(* Logix 5000 project; controller TFF vendor 1 type 14 code 107 rev 34.11; software revision 34.03; part 4 of 36 *)

        BufferEvents[140] := '07242026,07:35:58.6,700003,0.0,1.00000000', BufferEvents[141] := '07242026,07:35:58.7,1300205,2.00000000,4.00000000', BufferEvents[142] := '07242026,07:35:58.7,1300405,2.00000000,4.00000000', BufferEvents[143] := '07242026,07:35:58.7,1300505,2.00000000,4.00000000', BufferEvents[144] := '07242026,07:35:58.7,1300605,2.00000000,4.00000000', BufferEvents[145] := '07242026,07:35:58.7,1301105,2.00000000,4.00000000', BufferEvents[146] := '07242026,07:35:58.7,1301205,2.00000000,4.00000000', BufferEvents[147] := '07242026,07:35:58.7,1301305,2.00000000,4.00000000', BufferEvents[148] := '07242026,07:35:58.7,1301405,2.00000000,4.00000000', BufferEvents[149] := '07242026,07:35:58.8,2500101,0.0,1.00000000', BufferEvents[150] := '07242026,07:35:58.8,2500401,0.0,1.00000000', BufferEvents[151] := '07242026,07:35:58.8,2500801,1.00000000,0.0', BufferEvents[152] := '07242026,07:35:58.8,2501901,0.0,1.00000000', BufferEvents[153] := '07242026,08:54:51.3,305106,1.00000000,0.0', BufferEvents[154] := '07242026,08:55:09.5,305206,1.00000000,0.0', BufferEvents[155] := '07242026,08:56:06.6,305006,1.00000000,0.0', BufferEvents[156] := '07242026,09:12:34.6,300107,0.0,1.00000000', BufferEvents[157] := '07242026,09:14:51.8,700003,1.00000000,0.0', BufferEvents[158] := '07242026,09:14:51.8,300106,1.00000000,0.0', BufferEvents[159] := '07242026,09:14:51.8,300607,0.0,1.00000000', BufferEvents[160] := '07242026,09:14:51.8,300707,0.0,1.00000000', BufferEvents[161] := '07242026,09:14:51.9,305006,0.0,1.00000000', BufferEvents[162] := '07242026,09:14:51.9,305106,0.0,1.00000000', BufferEvents[163] := '07242026,09:14:51.9,305206,0.0,1.00000000', BufferEvents[164] := '07242026,09:14:51.9,1600003,1.00000000,0.0', BufferEvents[165] := '07242026,09:14:51.9,1300205,4.00000000,2.00000000', BufferEvents[166] := '07242026,09:14:51.9,1300405,4.00000000,2.00000000', BufferEvents[167] := '07242026,09:14:51.9,1300505,4.00000000,2.00000000', BufferEvents[168] := '07242026,09:14:51.9,1300605,4.00000000,2.00000000', BufferEvents[169] := '07242026,09:14:51.9,1301105,4.00000000,2.00000000', BufferEvents[170] := '07242026,09:14:51.9,1301205,4.00000000,2.00000000', BufferEvents[171] := '07242026,09:14:51.9,1301305,4.00000000,2.00000000', BufferEvents[172] := '07242026,09:14:51.9,1301405,4.00000000,2.00000000', BufferEvents[173] := '07242026,09:14:52.0,2500101,1.00000000,0.0', BufferEvents[174] := '07242026,09:14:52.0,2500401,1.00000000,0.0', BufferEvents[175] := '07242026,09:14:52.0,2500801,0.0,1.00000000', BufferEvents[176] := '07242026,09:14:52.0,2501901,1.00000000,0.0', BufferEvents[177] := '07242026,09:14:52.9,306806,1.00000000,0.0', BufferEvents[178] := '07242026,09:14:55.0,1600003,0.0,1.00000000', BufferEvents[179] := '07242026,09:14:56.8,305506,1.00000000,0.0', BufferEvents[180] := '07242026,09:14:56.8,305706,1.00000000,0.0', BufferEvents[181] := '07242026,09:14:56.8,306906,1.00000000,0.0', BufferEvents[182] := '07242026,09:14:56.8,307106,1.00000000,0.0', BufferEvents[183] := '07242026,09:14:56.8,307306,1.00000000,0.0', BufferEvents[184] := '07242026,09:14:56.8,307506,1.00000000,0.0', BufferEvents[185] := '07242026,09:15:07.7,300106,0.0,1.00000000', BufferEvents[186] := '07242026,09:15:07.7,306806,0.0,1.00000000', BufferEvents[187] := '07242026,09:15:07.7,300107,1.00000000,0.0', BufferEvents[188] := '07242026,09:15:07.7,300607,1.00000000,0.0', BufferEvents[189] := '07242026,09:15:07.7,300707,1.00000000,0.0', BufferEvents[190] := '07242026,09:15:07.8,300306,1.00000000,0.0', BufferEvents[191] := '07242026,09:15:09.7,300006,1.00000000,0.0', BufferEvents[192] := '07242026,09:19:10.3,305506,0.0,1.00000000', BufferEvents[193] := '07242026,09:19:10.3,305706,0.0,1.00000000', BufferEvents[194] := '07242026,09:19:10.3,307106,0.0,1.00000000', BufferEvents[195] := '07242026,09:19:10.3,307306,0.0,1.00000000', BufferEvents[196] := '07242026,09:19:10.3,307506,0.0,1.00000000', BufferEvents[197] := '07242026,09:19:10.3,1600003,1.00000000,0.0', BufferEvents[198] := '07242026,09:19:13.4,1600003,0.0,1.00000000', BufferEvents[199] := '07242026,09:19:17.6,300306,0.0,1.00000000',
        BufferEvents[200] := '07242026,09:19:18.6,300006,0.0,1.00000000', BufferEvents[201] := '07242026,09:19:35.6,306906,0.0,1.00000000', BufferEvents[202] := '07242026,09:19:36.6,300806,1.00000000,0.0', BufferEvents[203] := '07242026,09:19:36.6,300906,1.00000000,0.0', BufferEvents[204] := '07242026,09:19:37.7,301006,1.00000000,0.0', BufferEvents[205] := '07242026,09:19:39.5,300806,0.0,1.00000000', BufferEvents[206] := '07242026,09:19:39.5,300906,0.0,1.00000000', BufferEvents[207] := '07242026,09:19:39.5,301006,0.0,1.00000000', BufferEvents[208] := '07242026,09:19:39.5,1600003,1.00000000,0.0', BufferEvents[209] := '07242026,09:19:42.6,1600003,0.0,1.00000000', BufferEvents[210] := '07242026,10:57:37.4,700003,0.0,1.00000000', BufferEvents[211] := '07242026,10:57:37.5,1300205,2.00000000,4.00000000', BufferEvents[212] := '07242026,10:57:37.5,1300405,2.00000000,4.00000000', BufferEvents[213] := '07242026,10:57:37.5,1300505,2.00000000,4.00000000', BufferEvents[214] := '07242026,10:57:37.5,1300605,2.00000000,4.00000000', BufferEvents[215] := '07242026,10:57:37.5,1301105,2.00000000,4.00000000', BufferEvents[216] := '07242026,10:57:37.5,1301205,2.00000000,4.00000000', BufferEvents[217] := '07242026,10:57:37.5,1301305,2.00000000,4.00000000', BufferEvents[218] := '07242026,10:57:37.5,1301405,2.00000000,4.00000000', BufferEvents[219] := '07242026,10:57:37.6,2500101,0.0,1.00000000', BufferEvents[220] := '07242026,10:57:37.6,2500401,0.0,1.00000000', BufferEvents[221] := '07242026,10:57:37.6,2500801,1.00000000,0.0', BufferEvents[222] := '07242026,10:57:37.6,2501901,0.0,1.00000000', BufferEvents[223] := '07242026,10:57:44.5,900103,1.00000000,0.0', BufferEvents[224] := '07242026,10:57:48.7,500106,30.0000000,0.0', BufferEvents[225] := '07242026,10:57:54.2,900101,1.00000000,0.0', BufferEvents[226] := '07242026,10:57:54.2,500128,1.00000000,0.0', BufferEvents[227] := '07242026,10:58:25.0,500128,0.0,1.00000000', BufferEvents[228] := '07242026,10:58:25.0,500126,1.00000000,0.0', BufferEvents[229] := '07242026,11:03:15.0,900101,0.0,1.00000000', BufferEvents[230] := '07242026,11:03:15.0,500126,0.0,1.00000000', BufferEvents[231] := '07242026,11:03:21.9,500106,0.0,30.0000000', BufferEvents[232] := '07242026,11:03:46.9,900103,0.0,1.00000000', BufferEvents[233] := '07242026,11:05:12.4,1700011,0.0,1.00000000', BufferEvents[234] := '07242026,11:05:12.5,1700003,1.00000000,0.0', BufferEvents[235] := '07242026,11:05:13.6,2600007,1.00000000,0.0', BufferEvents[236] := '07242026,11:05:13.6,2600007,0.0,1.00000000', BufferEvents[237] := '07242026,11:05:13.8,700005,10.0000000,0.0', BufferEvents[238] := '07242026,11:05:13.9,700301,1.00000000,0.0', BufferEvents[239] := '07242026,11:05:13.9,700302,0.0,1.00000000', BufferEvents[240] := '07242026,11:05:14.1,1301205,4.00000000,2.00000000', BufferEvents[241] := '07242026,11:05:14.1,1301305,4.00000000,2.00000000', BufferEvents[242] := '07242026,11:05:14.2,2502801,1.00000000,0.0', BufferEvents[243] := '07242026,11:05:14.2,1301205,2.00000000,4.00000000', BufferEvents[244] := '07242026,11:05:14.3,2502801,0.0,1.00000000', BufferEvents[245] := '07242026,11:05:14.3,2300001,1.00000000,0.0', BufferEvents[246] := '07242026,11:05:14.3,1301305,2.00000000,4.00000000', BufferEvents[247] := '07242026,11:05:14.4,2300003,1.00000000,0.0', BufferEvents[248] := '07242026,11:05:14.5,800301,1.00000000,0.0', BufferEvents[249] := '07242026,11:05:15.4,2300001,0.0,1.00000000', BufferEvents[250] := '07242026,11:05:15.5,2300003,0.0,1.00000000', DefaultOnComplete := 1);   // CCP System Data
   CCPSystem_Storage : CCPSystem_Storage[6] := ([0].Download := 1, [0].TestAction := 1, [0].State := 3, [0].Language := 1, [0].EndPointer := 34, [0].Machine := 'Mobius FlexReady', [0].Created := '03/13/2018 4:36:30 AM', [0].Originator := 'Smart', [0].OperationName := 'c:\\millipore\\CCPRecipeFiles\\SmartXMO_00.02.opn', [0].ConfigFile := 'XMO4.cfg', [0].StateWatchDog.PRE := 300000, [1].Download := 1, [1].TestAction := 1, [1].State := 3, [1].Language := 1, [1].EndPointer := 1, [1].Machine := 'Mobius FlexReady', [1].Created := '08/06/2019 8:22:36 AM', [1].Originator := 'test', [1].ConfigFile := 'TF3S.cfg', [1].StateWatchDog.PRE := 300000, [2].Download := 1, [2].TestAction := 1, [2].State := 3, [2].Language := 1, [2].EndPointer := 5, [2].Machine := 'Mobius FlexReady', [2].Created := '02/20/2018 2:20:36 AM', [2].Originator := 'QSP', [2].ConfigFile := 'MASTER_CFG--XMO4.cfg', [2].StateWatchDog.PRE := 300000, [3].Download := 1, [3].OperationDownloadFlag := 1, [3].TestAction := 1, [3].State := 3, [3].Language := 1, [3].EndPointer := 9, [3].Machine := 'Mobius FlexReady', [3].Created := '01/18/2018 5:35:26 AM', [3].Originator := 'ccc', [3].OperationName := 'c:\\millipore\\CCPRecipeFiles\\Untitled2_00.02.opn', [3].ConfigFile := 'MASTER_CFG--XMO4.cfg', [3].StateWatchDog.PRE := 300000, [4].Download := 1, [4].TestAction := 1, [4].State := 3, [4].Language := 1, [4].EndPointer := 9, [4].Machine := 'Mobius FlexReady', [4].Created := '01/18/2018 5:35:26 AM', [4].Originator := 'ccc', [4].ConfigFile := 'MASTER_CFG--XMO4.cfg', [4].StateWatchDog.PRE := 300000, [5].Download := 1, [5].OperationDownloadFlag := 1, [5].TestAction := 1, [5].State := 3, [5].Language := 1, [5].EndPointer := 9, [5].Machine := 'Mobius FlexReady',
        [5].Created := '01/18/2018 5:35:26 AM', [5].Originator := 'ccc', [5].OperationName := 'c:\\millipore\\CCPRecipeFiles\\Untitled2_00.02.opn', [5].ConfigFile := 'MASTER_CFG--XMO4.cfg', [5].StateWatchDog.PRE := 300000);
   ChartMark : ChartMark := (Out := 1);   // Chart Mark
   Concentration : Concentration := (VCF := 1.0, CB := 15.9, Conc_Init := 15.9, Conc_Final := 30.0, Final_Conc_Volume_Reached := 1, Final_Conc_Volume_DownTimer.PRE := 10000, Final_Conc_Volume_UpTimer.PRE := 1000, Final_Conc_Volume_UpTimer.ACC := 1015, Final_Conc_Volume_UpTimer.EN := 1, Final_Conc_Volume_UpTimer.DN := 1, Final_Conc_Protein_DownTimer.PRE := 10000, Final_Conc_Protein_DownTimer.ACC := 10089, Final_Conc_Protein_DownTimer.EN := 1, Final_Conc_Protein_DownTimer.DN := 1, Final_Conc_Protein_UpTimer.PRE := 1000, LogConcTimer.PRE := 3000);
   ControlLoop : ControlLoop[20] := ([0].RampTimer.PRE := 3600000, [0].StableTimer.PRE := 5000, [0].PIDTimer.PRE := 250, [0].PIDTimer.ACC := 100, [0].PIDTimer.EN := 1, [0].PIDTimer.TT := 1, [0].PID.CTL := 25199488, [0].PID.MO := 1, [0].PID.PE := 1, [0].PID.INI := 1, [0].PID.DVPA := 1, [0].PID.PVLA := 1, [0].PID.PVHA := 1, [0].PID.SP := 66.66666, [0].PID.KP := 0.5, [0].PID.KI := 0.1, [0].PID.MAXS := 200.0, [0].PID.SO := 10.0, [0].PID.MAXO := 100.0, [0].PID.MINO := 10.0, [0].PID.UPD := 0.25, [0].PID.ERR := 66.66666, [0].PID.OUT := 10.0, [0].PID.MAXI := 200.0, [0].PID.TIE := 10.0, [0].PID.MAXCV := 100.0, [0].PID.MAXTIE := 100.0, [0].PID.DATA[0] := -6.666666, [0].PID.DATA[3] := 66.66666, [0].PID.DATA[4] := 66.66666, [0].PID.DATA[5] := 0.5, [0].PID.DATA[6] := 1.0, [0].PID.DATA[7] := 4.0, [0].PID.DATA[8] := 0.5, [0].PID.DATA[9] := 0.1, [0].PID.DATA[11] := 0.5, [0].PID.DATA[12] := 0.08333334, [0].PID.DATA[15] := 1.0, [0].PID.DATA[16] := 1.0, [1].Tag := 'FIC01', [1].Desc := 'Feed Pump Control Loop', [1].LoopCfg := 1, [1].ManualEGU := '%', [1].Auto1EGU := 'LPM', [1].Auto2EGU := 'Bar', [1].Manual := 1, [1].RampEnable := 1, [1].PIDEnable := 1, [1].ManualOSR := 1, [1].PVAuto2 := 3.9859235, [1].SPAuto := 10.0, [1].SPAuto1 := 10.0, [1].SPAuto2 := 1.0, [1].RangeMax := 100.0, [1].RampRate := 1.0, [1].RampRateSave := 1.0, [1].Deadband := 10.0, [1].DBLO := 9.0, [1].DBHI := 11.0, [1].RampTimer.PRE := 3600000,
        [1].StableTimer.PRE := 10000, [1].StableTime := 10, [1].PIDTimer.PRE := 250, [1].CycleTimer.PRE := 2000, [1].PID.CTL := -2080341120, [1].PID.EN := 1, [1].PID.SWM := 1, [1].PID.INI := 1, [1].PID.DVPA := 1, [1].PID.PVLA := 1, [1].PID.PVHA := 1, [1].PID.SP := 10.0, [1].PID.KP := 0.1, [1].PID.KI := 0.2, [1].PID.MAXS := 48.0, [1].PID.DB := 0.01, [1].PID.MAXO := 100.0, [1].PID.UPD := 0.25, [1].PID.ERR := 10.0, [1].PID.MAXI := 48.0, [1].PID.MAXCV := 100.0, [1].PID.MAXTIE := 48.0, [1].PID.DATA[0] := -2.0833333, [1].PID.DATA[3] := 10.0, [1].PID.DATA[4] := 10.0, [1].PID.DATA[5] := 2.0833333, [1].PID.DATA[6] := 1.0, [1].PID.DATA[7] := 4.0, [1].PID.DATA[8] := 0.1, [1].PID.DATA[9] := 0.2, [1].PID.DATA[11] := 0.1, [1].PID.DATA[12] := 0.2, [1].PID.DATA[15] := 1.0, [1].PID.DATA[16] := 2.0833333, [1].KP[0] := 100.0, [1].KP[1] := 100.0, [1].KI[0] := 200.0, [1].KI[1] := 200.0, [1].DB[0] := 0.01, [1].Auto1Cfg := 1, [1].Auto2Cfg := 1, [1].Auto1PVCfg := 42, [1].Auto2PVCfg := 40, [1].Auto1RangeMax := 48.0, [1].Auto2RangeMax := 87.0, [1].OutputAddress := 2, [2].Tag := 'LIC01', [2].Desc := 'Level Control Loop', [2].LoopCfg := 1, [2].ManualEGU := '%', [2].Auto1EGU := 'L', [2].Interlock := 1, [2].Manual := 1, [2].RampEnable := 1, [2].PIDEnable := 1, [2].ManualOSR := 1, [2].PVAuto2 := 2400.0, [2].SPAuto := 51.59, [2].SPAuto1 := 51.59, [2].RangeMax := 100.0,
        [2].RampRate := 5.0, [2].RampRateSave := 5.0, [2].Deadband := 15.0, [2].DBLO := 43.8515, [2].DBHI := 59.3285, [2].RampTimer.PRE := 3600000, [2].StableTimer.PRE := 10000, [2].StableTime := 10, [2].PIDTimer.PRE := 250, [2].CycleTimer.PRE := 2000, [2].PID.CTL := -2080341120, [2].PID.EN := 1, [2].PID.SWM := 1, [2].PID.INI := 1, [2].PID.DVPA := 1, [2].PID.PVLA := 1, [2].PID.PVHA := 1, [2].PID.SP := 51.59, [2].PID.KP := 5.0, [2].PID.KI := 10.0, [2].PID.MAXS := 200.0, [2].PID.DB := 0.001, [2].PID.MAXO := 100.0, [2].PID.UPD := 0.25, [2].PID.ERR := 51.59, [2].PID.MAXI := 200.0, [2].PID.MAXCV := 100.0, [2].PID.MAXTIE := 100.0, [2].PID.DATA[0] := -128.975, [2].PID.DATA[3] := 51.59, [2].PID.DATA[4] := 51.59, [2].PID.DATA[5] := 0.5, [2].PID.DATA[6] := 1.0, [2].PID.DATA[7] := 4.0, [2].PID.DATA[8] := 5.0, [2].PID.DATA[9] := 10.0, [2].PID.DATA[11] := 5.0, [2].PID.DATA[12] := 10.0, [2].PID.DATA[15] := 1.0, [2].PID.DATA[16] := 1.0, [2].KP[0] := 5000.0, [2].KP[1] := 5000.0, [2].KI[0] := 10000.0, [2].KI[1] := 10000.0, [2].DB[0] := 0.001, [2].DisOSR := 1, [2].Auto1Cfg := 1, [2].Auto1PVCfg := 44, [2].Auto1RangeMax := 200.0, [2].OutputAddress := 3, [3].Tag := 'Mixer', [3].LoopCfg := 1, [3].ManualEGU := '%', [3].Enable := 1, [3].Manual := 1, [3].Stable := 1, [3].Status := 3, [3].RampEnable := 1, [3].PIDEnable := 1, [3].ManualOSR := 1,
        [3].PV := -0.20576791, [3].PVAuto1 := -0.20576791, [3].PVAuto2 := 20.902039, [3].CV := 2.2879825, [3].SPAuto := 6.0, [3].SPAutoSave := -0.20576791, [3].SPAuto1 := 6.0, [3].SPAuto2 := 20.0, [3].RangeMax := 100.0, [3].RampRate := 2.0, [3].RampRateSave := 2.0, [3].Deadband := 20.0, [3].DBLO := 4.8, [3].DBHI := 7.2, [3].RampTimer.PRE := 3600000, [3].StableTimer.PRE := 10000, [3].StableTime := 10, [3].PIDTimer.PRE := 250, [3].CycleTimer.PRE := 2000, [3].PID.CTL := -2080341248, [3].PID.EN := 1, [3].PID.SWM := 1, [3].PID.INI := 1, [3].PID.DVPA := 1, [3].PID.PVLA := 1, [3].PID.SP := 6.0, [3].PID.KP := 0.04, [3].PID.KI := 0.04, [3].PID.BIAS := 30.796, [3].PID.MAXS := 87.0, [3].PID.DB := 0.02, [3].PID.SO := 2.2879825, [3].PID.MAXO := 100.0, [3].PID.UPD := 0.25, [3].PID.PV := -0.20576791, [3].PID.ERR := 6.205768, [3].PID.OUT := 2.2879825, [3].PID.MAXI := 87.0, [3].PID.TIE := 2.2879825, [3].PID.MAXCV := 100.0, [3].PID.MAXTIE := 100.0, [3].PID.DATA[0] := -28.793339, [3].PID.DATA[1] := 3.7842374, [3].PID.DATA[2] := -0.20576791, [3].PID.DATA[3] := 6.205768, [3].PID.DATA[4] := 6.0, [3].PID.DATA[5] := 1.1494253, [3].PID.DATA[6] := 1.0, [3].PID.DATA[7] := 4.0, [3].PID.DATA[8] := 0.04, [3].PID.DATA[9] := 0.04, [3].PID.DATA[11] := 0.04, [3].PID.DATA[12] := 0.04, [3].PID.DATA[15] := 1.0, [3].PID.DATA[16] := 1.0, [3].KP[0] := 40.0, [3].KP[1] := 40.0, [3].KI[0] := 40.0, [3].KI[1] := 40.0, [3].DB[0] := 0.02,
        [3].DB[1] := 0.02, [3].Auto1Cfg := 1, [3].Auto2Cfg := 1, [3].Auto1PVCfg := 6, [3].Auto2PVCfg := 41, [3].Auto1RangeMax := 87.0, [3].Auto2RangeMax := 87.0, [4].Tag := 'PC001', [4].Desc := 'Retentate Control Valve', [4].ManualEGU := '%', [4].Auto1EGU := 'Bar', [4].Auto2EGU := 'Bar', [4].Enable := 1, [4].Status := 3, [4].PIDEnable := 1, [4].PV := -0.09876543, [4].PVAuto1 := -1.4998856, [4].CV := 2.2879825, [4].SPAutoSave := 101.99314, [4].RangeMax := 100.0, [4].RampRate := 2.4, [4].RampRateSave := 2.4, [4].Deadband := 10.0, [4].RampTimer.PRE := 3600000, [4].StableTimer.PRE := 5000, [4].StableTime := 5, [4].PIDTimer.PRE := 250, [4].CycleTimer.PRE := 2000, [4].PID.CTL := -2145350912, [4].PID.EN := 1, [4].PID.NOBC := 1, [4].PID.INI := 1, [4].PID.EWD := 1, [4].PID.DVPA := 1, [4].PID.PVLA := 1, [4].PID.KP := 0.2, [4].PID.KI := 0.08, [4].PID.KD := 0.01, [4].PID.MAXS := 100.0, [4].PID.DB := 0.3, [4].PID.SO := 2.2879825, [4].PID.MAXO := 100.0, [4].PID.UPD := 0.005, [4].PID.PV := -0.09876543, [4].PID.ERR := 0.09876543, [4].PID.OUT := 2.2879825, [4].PID.MAXI := 100.0, [4].PID.TIE := 0.05587259, [4].PID.MAXCV := 100.0, [4].PID.MAXTIE := 4095.0, [4].PID.DATA[0] := 2.281907, [4].PID.DATA[1] := 1.5168943, [4].PID.DATA[2] := -0.09876543, [4].PID.DATA[3] := 0.09876543, [4].PID.DATA[5] := 1.0, [4].PID.DATA[6] := 1.0, [4].PID.DATA[7] := 0.089999996, [4].PID.DATA[8] := 0.2, [4].PID.DATA[9] := 0.08, [4].PID.DATA[10] := 0.01,
        [4].PID.DATA[11] := 0.2, [4].PID.DATA[12] := 0.08, [4].PID.DATA[13] := 0.01, [4].PID.DATA[15] := 1.0, [4].PID.DATA[16] := 0.024420025, [4].KP[0] := 40.0, [4].KP[1] := 40.0, [4].KI[0] := 1.0, [4].KI[1] := 40.0, [4].DB[0] := 0.02, [5].LoopCfg := 1, [5].ManualEGU := '%', [5].Enable := 1, [5].Manual := 1, [5].Stable := 1, [5].Status := 3, [5].RampEnable := 1, [5].PIDEnable := 1, [5].ManualOSR := 1, [5].PVAuto2 := 0.23729686, [5].CV := 86.54368, [5].SPAuto2 := 11.0, [5].SPManual := 100.0, [5].SPManualSave := 100.0, [5].RangeMax := 100.0, [5].RampRate := 5.0, [5].RampRateSave := 5.0, [5].RampStart := 100.0, [5].Deadband := 10.0, [5].RampTimer.PRE := 3600000, [5].StableTimer.PRE := 10000, [5].StableTime := 10, [5].PIDTimer.PRE := 250, [5].CycleTimer.PRE := 2000, [5].PID.CTL := -2080340096, [5].PID.EN := 1, [5].PID.SWM := 1, [5].PID.INI := 1, [5].PID.DVNA := 1, [5].PID.DVPA := 1, [5].PID.PVLA := 1, [5].PID.PVHA := 1, [5].PID.KP := 0.25, [5].PID.KI := 0.1, [5].PID.KD := 0.1, [5].PID.BIAS := -847.4798, [5].PID.MAXS := 20.0, [5].PID.DB := 0.02, [5].PID.SO := 86.54368, [5].PID.MAXO := 100.0, [5].PID.UPD := 0.25, [5].PID.OUT := 86.54368, [5].PID.MAXI := 20.0, [5].PID.TIE := 86.47018, [5].PID.MAXCV := 100.0, [5].PID.MAXTIE := 100.0, [5].PID.DATA[0] := 934.0235, [5].PID.DATA[5] := 5.0, [5].PID.DATA[6] := 1.0, [5].PID.DATA[7] := 4.1,
        [5].PID.DATA[8] := 0.25, [5].PID.DATA[9] := 0.1, [5].PID.DATA[10] := 0.1, [5].PID.DATA[11] := 0.25, [5].PID.DATA[12] := 0.1, [5].PID.DATA[13] := 0.1, [5].PID.DATA[15] := 1.0, [5].PID.DATA[16] := 1.0, [5].KP[0] := 250.0, [5].KP[1] := 250.0, [5].KI[0] := 100.0, [5].KI[1] := 100.0, [5].KD[0] := 100.0, [5].KD[1] := 100.0, [5].DB[0] := 0.02, [5].DB[1] := 0.02, [5].Auto1Cfg := 1, [5].Auto2Cfg := 1, [5].Auto1PVCfg := 2, [5].Auto2PVCfg := 41, [5].Auto1RangeMax := 20.0, [5].Auto2RangeMax := 87.0, [5].OutputAddress := 1, [6].Tag := 'PC101', [6].Desc := 'Filtrate Control Valve', [6].AutoEGU := 'Bar', [6].Auto1EGU := 'Bar', [6].Enable := 1, [6].Stable := 1, [6].DBOK := 1, [6].Status := 3, [6].PIDEnable := 1, [6].PV := 99.47403, [6].PVAuto1 := -6.249523, [6].CV := 86.51909, [6].SPAuto := 100.0, [6].SPAutoSave := 38.696636, [6].RangeMax := 100.0, [6].RampRate := 6.0, [6].RampRateSave := 6.0, [6].Deadband := 10.0, [6].DBLO := 90.0, [6].DBHI := 110.0, [6].RampTimer.PRE := 3600000, [6].StableTimer.PRE := 5000, [6].StableTime := 5, [6].PIDTimer.PRE := 250, [6].PIDTimer.EN := 1, [6].PIDTimer.TT := 1, [6].CycleTimer.PRE := 2000, [6].PID.CTL := 2130560, [6].PID.NOBC := 1, [6].PID.INI := 1, [6].PID.DVPA := 1, [6].PID.PVHA := 1, [6].PID.SP := 100.0, [6].PID.KP := 0.3, [6].PID.KI := 0.08, [6].PID.KD := 0.01, [6].PID.MAXS := 100.0,
        [6].PID.DB := 0.3, [6].PID.SO := 86.51909, [6].PID.MAXO := 100.0, [6].PID.UPD := 0.005, [6].PID.PV := 99.47403, [6].PID.ERR := 0.52597046, [6].PID.OUT := 86.51909, [6].PID.MAXI := 100.0, [6].PID.TIE := 2.113094, [6].PID.MAXCV := 100.0, [6].PID.MAXTIE := 4095.0, [6].PID.DATA[0] := 86.32628, [6].PID.DATA[1] := -1591.6195, [6].PID.DATA[2] := 99.47403, [6].PID.DATA[3] := 0.52597046, [6].PID.DATA[4] := 100.0, [6].PID.DATA[5] := 1.0, [6].PID.DATA[6] := 1.0, [6].PID.DATA[7] := 0.089999996, [6].PID.DATA[8] := 0.3, [6].PID.DATA[9] := 0.08, [6].PID.DATA[10] := 0.01, [6].PID.DATA[11] := 0.3, [6].PID.DATA[12] := 0.08, [6].PID.DATA[13] := 0.01, [6].PID.DATA[15] := 1.0, [6].PID.DATA[16] := 0.024420025, [6].KP[0] := 100.0, [6].KP[1] := 250.0, [6].KI[0] := 5.0, [6].KI[1] := 20.0, [6].DB[0] := 0.02, [6].OutputAddress := 1, [7].StableTimer.PRE := 200, [7].PIDTimer.PRE := 250, [7].PIDTimer.EN := 1, [7].PIDTimer.TT := 1, [7].CycleTimer.PRE := 10000, [7].PID.CTL := 16810880, [7].PID.MO := 1, [7].PID.INI := 1, [7].PID.DVPA := 1, [7].PID.PVLA := 1, [7].PID.PVHA := 1, [7].PID.SP := 10.0, [7].PID.KP := 2.0, [7].PID.KI := 0.2, [7].PID.KD := 0.3, [7].PID.BIAS := 50.0, [7].PID.DB := 0.01, [7].PID.SO := 80.0, [7].PID.MAXO := 100.0, [7].PID.UPD := 0.25, [7].PID.ERR := 10.0, [7].PID.OUT := 80.0, [7].PID.TIE := 80.0, [7].PID.MAXCV := 100.0, [7].PID.MAXTIE := 100.0, [7].PID.DATA[0] := 29.5116, [7].PID.DATA[3] := 10.0,
        [7].PID.DATA[4] := 10.0, [7].PID.DATA[5] := 0.02442002, [7].PID.DATA[6] := 1.0, [7].PID.DATA[7] := 4.3, [7].PID.DATA[8] := 2.0, [7].PID.DATA[9] := 0.2, [7].PID.DATA[10] := 0.3, [7].PID.DATA[11] := 2.0, [7].PID.DATA[12] := 0.2, [7].PID.DATA[13] := 0.3, [7].PID.DATA[15] := 1.0, [7].PID.DATA[16] := 1.0, [8].StableTimer.PRE := 15000, [8].PIDTimer.PRE := 250, [8].CycleTimer.PRE := 20000, [8].PID.CTL := 33555584, [8].PID.CA := 1, [8].PID.DVNA := 1, [8].PID.PVHA := 1, [8].PID.SP := 27.0, [8].PID.KP := 1.0, [8].PID.KI := 0.1, [8].PID.MAXS := 100.0, [8].PID.MAXO := 100.0, [8].PID.UPD := 0.25, [8].PID.PV := 18.2328, [8].PID.ERR := -8.767202, [8].PID.MAXI := 100.0, [8].PID.MAXCV := 100.0, [8].PID.MAXTIE := 100.0, [8].PID.DATA[0] := 8.767202, [8].PID.DATA[1] := 291.7248, [8].PID.DATA[2] := 18.2328, [8].PID.DATA[3] := -8.767202, [8].PID.DATA[4] := 27.0, [8].PID.DATA[5] := 1.0, [8].PID.DATA[6] := 1.0, [8].PID.DATA[7] := 4.0, [8].PID.DATA[8] := 1.0, [8].PID.DATA[9] := 0.1, [8].PID.DATA[11] := 1.0, [8].PID.DATA[12] := 0.1, [8].PID.DATA[15] := 1.0, [8].PID.DATA[16] := 1.0, [11].RampTimer.PRE := 100000, [11].StableTimer.PRE := 200, [11].PIDTimer.PRE := 250, [11].PIDTimer.ACC := 230, [11].PIDTimer.EN := 1, [11].PIDTimer.TT := 1, [11].PID.CTL := 67142528, [11].PID.SWM := 1, [11].PID.INI := 1, [11].PID.DVPA := 1, [11].PID.PVLA := 1, [11].PID.PVHA := 1, [11].PID.SP := 0.2, [11].PID.KP := 0.1, [11].PID.KI := 0.1, [11].PID.BIAS := 23.09767,
        [11].PID.DB := 0.001, [11].PID.MAXO := 100.0, [11].PID.UPD := 0.25, [11].PID.ERR := 0.2, [11].PID.MAXCV := 100.0, [11].PID.MAXTIE := 100.0, [11].PID.DATA[0] := -23.09816, [11].PID.DATA[3] := 0.2, [11].PID.DATA[4] := 0.2, [11].PID.DATA[5] := 0.02442002, [11].PID.DATA[6] := 1.0, [11].PID.DATA[7] := 4.0, [11].PID.DATA[8] := 0.1, [11].PID.DATA[9] := 0.1, [11].PID.DATA[11] := 0.1, [11].PID.DATA[12] := 0.1, [11].PID.DATA[15] := 1.0, [11].PID.DATA[16] := 1.0, [13].RampTimer.PRE := 3600000, [13].StableTimer.PRE := 2000, [13].PIDTimer.PRE := 10000, [13].PIDTimer.EN := 1, [13].PIDTimer.TT := 1, [13].PID.CTL := 305173120, [13].PID.PVT := 1, [13].PID.CA := 1, [13].PID.NOBC := 1, [13].PID.NOZC := 1, [13].PID.INI := 1, [13].PID.OLH := 1, [13].PID.DVPA := 1, [13].PID.PVHA := 1, [13].PID.KP := 0.2, [13].PID.KI := 0.08, [13].PID.MAXS := 100.0, [13].PID.DB := 1.0, [13].PID.SO := 100.0, [13].PID.MAXO := 100.0, [13].PID.UPD := 0.01, [13].PID.PV := 43.92523, [13].PID.ERR := 43.92523, [13].PID.OUT := 100.0, [13].PID.MAXI := 100.0, [13].PID.TIE := 2.442003, [13].PID.MAXCV := 100.0, [13].PID.MAXTIE := 4095.0, [13].PID.DATA[0] := 100.0, [13].PID.DATA[1] := 702.8037, [13].PID.DATA[2] := 43.92523, [13].PID.DATA[3] := 43.92523, [13].PID.DATA[5] := 1.0, [13].PID.DATA[6] := 1.0, [13].PID.DATA[7] := 0.16, [13].PID.DATA[8] := 0.2, [13].PID.DATA[9] := 0.08, [13].PID.DATA[11] := 0.2, [13].PID.DATA[12] := 0.08, [13].PID.DATA[15] := 1.0, [13].PID.DATA[16] := 0.02442002);   // Control Loop Array
        [2]   // LIC001 Level Control Loop
        [3]   // PCV001 Control Loop
        [5]   // PCV101 Control Loop
        [4]   // PCV001 5ms Control Loop
        [6]   // PCV101 5ms Control Loop
        [1]   // FIC001 Feed Pump Control Loop
   ControlLoop_FeedBagLevel : ALIAS FOR ControlLoop[2];   // Feed Bag Level Control Loop
   ControlLoop_FeedBagLevelAlarm : ALIAS FOR AlarmDeviation[2];   // Feed Bag Level Control Loop Deviation Alarm
   ControlLoop_FeedPump : ALIAS FOR ControlLoop[1];   // Feed Pump Control Loop
   ControlLoop_FeedPumpAlarm : ALIAS FOR AlarmDeviation[1];   // Feed Pump Control Loop Deviation Alarm
   ControlLoop_PCV001 : ALIAS FOR ControlLoop[3];   // PCV001 Control Loop
   ControlLoop_PCV001_5ms : ALIAS FOR ControlLoop[4];   // PCV001 Control Loop
   ControlLoop_PCV001_CV : REAL;   // Control Value
   ControlLoop_PCV001_RAMP_OUT : REAL;   // Ramp Output
   ControlLoop_PCV001Alarm : ALIAS FOR AlarmDeviation[3];   // PCV001 Control Loop Deviation Alarm
   ControlLoop_PCV101 : ALIAS FOR ControlLoop[5];   // PCV101 Control Loop
   ControlLoop_PCV101_5ms : ALIAS FOR ControlLoop[6];   // PCV101 Control Loop
   ControlLoop_PCV101_CV : REAL := 100.0;   // Control Value
   ControlLoop_PCV101_RAMP_OUT : REAL := 100.0;   // Ramp Output
   ControlLoop_PCV101Alarm : ALIAS FOR AlarmDeviation[5];   // PCV101 Control Loop Deviation Alarm
   ControlLoop_Storage : ControlLoop[6,20] := ([0,0].RampTimer.PRE := 3600000, [0,0].StableTimer.PRE := 5000, [0,0].PIDTimer.PRE := 250, [0,0].PIDTimer.ACC := 100, [0,0].PIDTimer.EN := 1, [0,0].PIDTimer.TT := 1, [0,0].PID.CTL := 25199488, [0,0].PID.MO := 1, [0,0].PID.PE := 1, [0,0].PID.INI := 1, [0,0].PID.DVPA := 1, [0,0].PID.PVLA := 1, [0,0].PID.PVHA := 1, [0,0].PID.SP := 66.66666, [0,0].PID.KP := 0.5, [0,0].PID.KI := 0.1, [0,0].PID.MAXS := 200.0, [0,0].PID.SO := 10.0, [0,0].PID.MAXO := 100.0, [0,0].PID.MINO := 10.0, [0,0].PID.UPD := 0.25, [0,0].PID.ERR := 66.66666, [0,0].PID.OUT := 10.0, [0,0].PID.MAXI := 200.0, [0,0].PID.TIE := 10.0, [0,0].PID.MAXCV := 100.0, [0,0].PID.MAXTIE := 100.0, [0,0].PID.DATA[0] := -6.666666, [0,0].PID.DATA[3] := 66.66666, [0,0].PID.DATA[4] := 66.66666, [0,0].PID.DATA[5] := 0.5, [0,0].PID.DATA[6] := 1.0, [0,0].PID.DATA[7] := 4.0, [0,0].PID.DATA[8] := 0.5, [0,0].PID.DATA[9] := 0.1, [0,0].PID.DATA[11] := 0.5, [0,0].PID.DATA[12] := 0.08333334, [0,0].PID.DATA[15] := 1.0, [0,0].PID.DATA[16] := 1.0, [0,1].Tag := 'FIC01', [0,1].Desc := 'Prim. Feed Pump Control', [0,1].LoopCfg := 1, [0,1].ManualEGU := '%', [0,1].Auto1EGU := 'LPM', [0,1].Auto2EGU := 'cm/h', [0,1].Manual := 1, [0,1].DBOK := 1, [0,1].RampEnable := 1, [0,1].PIDEnable := 1, [0,1].ManualOSR := 1, [0,1].RangeMax := 100.0, [0,1].RampRate := 5.0, [0,1].RampRateSave := 5.0, [0,1].Deadband := 5.0, [0,1].RampTimer.PRE := 3600000, [0,1].StableTimer.PRE := 10000, [0,1].StableTime := 10, [0,1].PIDTimer.PRE := 250, [0,1].CycleTimer.PRE := 2000, [0,1].PID.CTL := -2080340096,
        [0,1].PID.EN := 1, [0,1].PID.SWM := 1, [0,1].PID.INI := 1, [0,1].PID.DVNA := 1, [0,1].PID.DVPA := 1, [0,1].PID.PVLA := 1, [0,1].PID.PVHA := 1, [0,1].PID.KP := 0.7, [0,1].PID.KI := 1.4, [0,1].PID.KD := 0.013, [0,1].PID.MAXS := 22.0, [0,1].PID.DB := 0.001, [0,1].PID.MAXO := 100.0, [0,1].PID.UPD := 0.25, [0,1].PID.MAXI := 22.0, [0,1].PID.MAXCV := 100.0, [0,1].PID.MAXTIE := 22.0, [0,1].PID.DATA[5] := 4.5454545, [0,1].PID.DATA[6] := 1.0, [0,1].PID.DATA[7] := 4.013, [0,1].PID.DATA[8] := 0.7, [0,1].PID.DATA[9] := 1.4, [0,1].PID.DATA[10] := 0.013, [0,1].PID.DATA[11] := 0.7, [0,1].PID.DATA[12] := 1.4, [0,1].PID.DATA[13] := 0.013, [0,1].PID.DATA[15] := 1.0, [0,1].PID.DATA[16] := 4.5454545, [0,1].KP[0] := 700.0, [0,1].KI[0] := 1400.0, [0,1].KD[0] := 13.0, [0,1].Auto1Cfg := 1, [0,1].Auto2Cfg := 1, [0,1].Auto1PVCfg := 10, [0,1].Auto2PVCfg := 42, [0,1].Auto1RangeMax := 22.0, [0,1].Auto2RangeMax := 9999.0, [0,2].Tag := 'FIC02', [0,2].Desc := 'Sec. Feed Pump Control', [0,2].LoopCfg := 1, [0,2].ManualEGU := '%', [0,2].Auto1EGU := 'LPM', [0,2].Auto2EGU := 'cm/h', [0,2].Interlock := 1, [0,2].Manual := 1, [0,2].DBOK := 1, [0,2].RampEnable := 1, [0,2].PIDEnable := 1, [0,2].ManualOSR := 1, [0,2].RangeMax := 100.0, [0,2].RampRate := 5.0, [0,2].RampRateSave := 5.0, [0,2].Deadband := 5.0, [0,2].RampTimer.PRE := 3600000, [0,2].StableTimer.PRE := 10000, [0,2].StableTime := 10, [0,2].PIDTimer.PRE := 250, [0,2].CycleTimer.PRE := 2000, [0,2].PID.CTL := -2080340096, [0,2].PID.EN := 1,
        [0,2].PID.SWM := 1, [0,2].PID.INI := 1, [0,2].PID.DVNA := 1, [0,2].PID.DVPA := 1, [0,2].PID.PVLA := 1, [0,2].PID.PVHA := 1, [0,2].PID.KP := 0.7, [0,2].PID.KI := 1.4, [0,2].PID.KD := 0.013, [0,2].PID.MAXS := 22.0, [0,2].PID.DB := 0.001, [0,2].PID.MAXO := 100.0, [0,2].PID.UPD := 0.25, [0,2].PID.MAXI := 22.0, [0,2].PID.MAXCV := 100.0, [0,2].PID.MAXTIE := 100.0, [0,2].PID.DATA[5] := 4.5454545, [0,2].PID.DATA[6] := 1.0, [0,2].PID.DATA[7] := 4.013, [0,2].PID.DATA[8] := 0.7, [0,2].PID.DATA[9] := 1.4, [0,2].PID.DATA[10] := 0.013, [0,2].PID.DATA[11] := 0.7, [0,2].PID.DATA[12] := 1.4, [0,2].PID.DATA[13] := 0.013, [0,2].PID.DATA[15] := 1.0, [0,2].PID.DATA[16] := 1.0, [0,2].KP[0] := 700.0, [0,2].KI[0] := 1400.0, [0,2].KD[0] := 13.0, [0,2].DisOSR := 1, [0,2].Auto1Cfg := 1, [0,2].Auto2Cfg := 1, [0,2].Auto1PVCfg := 12, [0,2].Auto2PVCfg := 43, [0,2].Auto1RangeMax := 22.0, [0,2].Auto2RangeMax := 9999.0, [0,2].OutputAddress := 1, [0,3].Tag := 'PCV12', [0,3].Desc := 'Post Column PCV012 Control', [0,3].LoopCfg := 1, [0,3].ManualEGU := '%', [0,3].Enable := 1, [0,3].Manual := 1, [0,3].Stable := 1, [0,3].DBOK := 1, [0,3].Status := 3, [0,3].RampEnable := 1, [0,3].PIDEnable := 1, [0,3].ManualOSR := 1, [0,3].RangeMax := 100.0, [0,3].RampRate := 5.0, [0,3].RampRateSave := 5.0, [0,3].RampStart := 20.0, [0,3].RampTimer.PRE := 3600000, [0,3].StableTimer.PRE := 2300, [0,3].StableTimer.ACC := 2354, [0,3].StableTimer.EN := 1, [0,3].StableTimer.DN := 1, [0,3].PIDTimer.PRE := 250,
        [0,3].CycleTimer.PRE := 2000, [0,3].PID.CTL := -1946122368, [0,3].PID.EN := 1, [0,3].PID.DOE := 1, [0,3].PID.SWM := 1, [0,3].PID.INI := 1, [0,3].PID.DVNA := 1, [0,3].PID.DVPA := 1, [0,3].PID.PVLA := 1, [0,3].PID.PVHA := 1, [0,3].PID.KP := 0.001, [0,3].PID.KI := 0.001, [0,3].PID.BIAS := 30.796, [0,3].PID.MAXS := 4095.0, [0,3].PID.MAXO := 100.0, [0,3].PID.UPD := 0.01, [0,3].PID.MAXI := 4095.0, [0,3].PID.MAXCV := 100.0, [0,3].PID.MAXTIE := 100.0, [0,3].PID.DATA[0] := -30.796, [0,3].PID.DATA[5] := 0.024420025, [0,3].PID.DATA[6] := 1.0, [0,3].PID.DATA[7] := 0.16, [0,3].PID.DATA[8] := 0.001, [0,3].PID.DATA[9] := 0.001, [0,3].PID.DATA[11] := 0.001, [0,3].PID.DATA[12] := 0.001, [0,3].PID.DATA[15] := 1.0, [0,3].PID.DATA[16] := 1.0, [0,3].OutputAddress := 2, [0,4].Tag := 'PCV10', [0,4].Desc := 'Line Pump1 PCV010 Control', [0,4].ManualEGU := '%', [0,4].Manual := 1, [0,4].Status := 3, [0,4].RampEnable := 1, [0,4].PIDEnable := 1, [0,4].RangeMax := 100.0, [0,4].RampRate := 0.5, [0,4].RampRateSave := 0.5, [0,4].RampStart := 3.443, [0,4].RampTimer.PRE := 3600000, [0,4].StableTimer.PRE := 5000, [0,4].PIDTimer.PRE := 250, [0,4].CycleTimer.PRE := 2000, [0,4].PID.CTL := 35652992, [0,4].PID.CA := 1, [0,4].PID.NOBC := 1, [0,4].PID.DVNA := 1, [0,4].PID.PVLA := 1, [0,4].PID.PVHA := 1, [0,4].PID.SP := 19.6, [0,4].PID.KP := 0.1, [0,4].PID.KI := 0.3, [0,4].PID.MAXS := 150.0, [0,4].PID.MAXO := 100.0, [0,4].PID.UPD := 0.25, [0,4].PID.ERR := -19.6, [0,4].PID.MAXI := 150.0, [0,4].PID.MAXCV := 100.0,
        [0,4].PID.MAXTIE := 100.0, [0,4].PID.DATA[0] := 1.3066667, [0,4].PID.DATA[3] := -19.6, [0,4].PID.DATA[4] := 19.6, [0,4].PID.DATA[5] := 0.6666667, [0,4].PID.DATA[6] := 1.0, [0,4].PID.DATA[7] := 4.0, [0,4].PID.DATA[8] := 0.1, [0,4].PID.DATA[9] := 0.3, [0,4].PID.DATA[11] := 0.1, [0,4].PID.DATA[12] := 0.3, [0,4].PID.DATA[15] := 1.0, [0,4].PID.DATA[16] := 1.0, [0,4].OutputAddress := 2, [0,5].Tag := 'PCV11', [0,5].Desc := 'Line Pump2 PCV011 Control', [0,5].ManualEGU := '%', [0,5].Manual := 1, [0,5].Status := 3, [0,5].RampEnable := 1, [0,5].PIDEnable := 1, [0,5].RangeMax := 100.0, [0,5].RampRate := 0.5, [0,5].RampRateSave := 0.5, [0,5].RampStart := 4.417, [0,5].RampTimer.PRE := 3600000, [0,5].StableTimer.PRE := 1500, [0,5].PIDTimer.PRE := 250, [0,5].CycleTimer.PRE := 2000, [0,5].PID.CTL := 134218624, [0,5].PID.DOE := 1, [0,5].PID.DVPA := 1, [0,5].PID.PVLA := 1, [0,5].PID.PVHA := 1, [0,5].PID.SP := 350.0, [0,5].PID.KP := 40.0, [0,5].PID.KI := 0.5, [0,5].PID.BIAS := -847.4798, [0,5].PID.MAXS := 550.0, [0,5].PID.MAXO := 100.0, [0,5].PID.UPD := 0.25, [0,5].PID.ERR := 350.0, [0,5].PID.MAXI := 550.0, [0,5].PID.MAXCV := 100.0, [0,5].PID.MAXTIE := 100.0, [0,5].PID.DATA[0] := -1697.9749, [0,5].PID.DATA[1] := 1018.1818, [0,5].PID.DATA[3] := 350.0, [0,5].PID.DATA[4] := 350.0, [0,5].PID.DATA[5] := 0.18181819, [0,5].PID.DATA[6] := 1.0, [0,5].PID.DATA[7] := 4.0, [0,5].PID.DATA[8] := 40.0, [0,5].PID.DATA[9] := 0.5, [0,5].PID.DATA[11] := 40.0, [0,5].PID.DATA[12] := 0.5, [0,5].PID.DATA[15] := 1.0, [0,5].PID.DATA[16] := 1.0, [0,5].OutputAddress := 3, [0,6].StableTimer.PRE := 15000,
        [0,6].PIDTimer.EN := 1, [0,6].PIDTimer.TT := 1, [0,6].CycleTimer.PRE := 5000, [0,6].PID.CTL := 16810624, [0,6].PID.MO := 1, [0,6].PID.INI := 1, [0,6].PID.DVPA := 1, [0,6].PID.PVHA := 1, [0,6].PID.SP := 10.0, [0,6].PID.KP := 0.3, [0,6].PID.KI := 0.3, [0,6].PID.MAXS := 200.0, [0,6].PID.SO := 3.074094, [0,6].PID.MAXO := 100.0, [0,6].PID.UPD := 0.25, [0,6].PID.PV := 1.488363, [0,6].PID.ERR := 8.511638, [0,6].PID.OUT := 3.074094, [0,6].PID.MAXI := 200.0, [0,6].PID.TIE := 3.074094, [0,6].PID.MAXCV := 200.0, [0,6].PID.MAXTIE := 200.0, [0,6].PID.DATA[0] := 1.797348, [0,6].PID.DATA[1] := -11.9069, [0,6].PID.DATA[2] := 1.488363, [0,6].PID.DATA[3] := 8.511638, [0,6].PID.DATA[4] := 10.0, [0,6].PID.DATA[5] := 0.5, [0,6].PID.DATA[6] := 1.0, [0,6].PID.DATA[7] := 4.0, [0,6].PID.DATA[8] := 0.3, [0,6].PID.DATA[9] := 0.3, [0,6].PID.DATA[11] := 0.3, [0,6].PID.DATA[12] := 0.3, [0,6].PID.DATA[15] := 2.0, [0,6].PID.DATA[16] := 0.5, [0,7].StableTimer.PRE := 200, [0,7].PIDTimer.PRE := 250, [0,7].PIDTimer.EN := 1, [0,7].PIDTimer.TT := 1, [0,7].CycleTimer.PRE := 10000, [0,7].PID.CTL := 16810880, [0,7].PID.MO := 1, [0,7].PID.INI := 1, [0,7].PID.DVPA := 1, [0,7].PID.PVLA := 1, [0,7].PID.PVHA := 1, [0,7].PID.SP := 10.0, [0,7].PID.KP := 2.0, [0,7].PID.KI := 0.2, [0,7].PID.KD := 0.3, [0,7].PID.BIAS := 50.0, [0,7].PID.DB := 0.01, [0,7].PID.SO := 80.0, [0,7].PID.MAXO := 100.0, [0,7].PID.UPD := 0.25, [0,7].PID.ERR := 10.0, [0,7].PID.OUT := 80.0, [0,7].PID.TIE := 80.0, [0,7].PID.MAXCV := 100.0,
        [0,7].PID.MAXTIE := 100.0, [0,7].PID.DATA[0] := 29.511597, [0,7].PID.DATA[3] := 10.0, [0,7].PID.DATA[4] := 10.0, [0,7].PID.DATA[5] := 0.024420025, [0,7].PID.DATA[6] := 1.0, [0,7].PID.DATA[7] := 4.3, [0,7].PID.DATA[8] := 2.0, [0,7].PID.DATA[9] := 0.2, [0,7].PID.DATA[10] := 0.3, [0,7].PID.DATA[11] := 2.0, [0,7].PID.DATA[12] := 0.2, [0,7].PID.DATA[13] := 0.3, [0,7].PID.DATA[15] := 1.0, [0,7].PID.DATA[16] := 1.0, [0,8].StableTimer.PRE := 15000, [0,8].PIDTimer.PRE := 250, [0,8].CycleTimer.PRE := 20000, [0,8].PID.CTL := 33555584, [0,8].PID.CA := 1, [0,8].PID.DVNA := 1, [0,8].PID.PVHA := 1, [0,8].PID.SP := 27.0, [0,8].PID.KP := 1.0, [0,8].PID.KI := 0.1, [0,8].PID.MAXS := 100.0, [0,8].PID.MAXO := 100.0, [0,8].PID.UPD := 0.25, [0,8].PID.PV := 18.2328, [0,8].PID.ERR := -8.767202, [0,8].PID.MAXI := 100.0, [0,8].PID.MAXCV := 100.0, [0,8].PID.MAXTIE := 100.0, [0,8].PID.DATA[0] := 8.767202, [0,8].PID.DATA[1] := 291.7248, [0,8].PID.DATA[2] := 18.2328, [0,8].PID.DATA[3] := -8.767202, [0,8].PID.DATA[4] := 27.0, [0,8].PID.DATA[5] := 1.0, [0,8].PID.DATA[6] := 1.0, [0,8].PID.DATA[7] := 4.0, [0,8].PID.DATA[8] := 1.0, [0,8].PID.DATA[9] := 0.1, [0,8].PID.DATA[11] := 1.0, [0,8].PID.DATA[12] := 0.1, [0,8].PID.DATA[15] := 1.0, [0,8].PID.DATA[16] := 1.0, [0,11].RampTimer.PRE := 100000, [0,11].StableTimer.PRE := 200, [0,11].PIDTimer.PRE := 250, [0,11].PIDTimer.ACC := 230, [0,11].PIDTimer.EN := 1, [0,11].PIDTimer.TT := 1, [0,11].PID.CTL := 67142528, [0,11].PID.SWM := 1, [0,11].PID.INI := 1, [0,11].PID.DVPA := 1, [0,11].PID.PVLA := 1, [0,11].PID.PVHA := 1, [0,11].PID.SP := 0.20000005,
        [0,11].PID.KP := 0.1, [0,11].PID.KI := 0.1, [0,11].PID.BIAS := 23.09767, [0,11].PID.DB := 0.001, [0,11].PID.MAXO := 100.0, [0,11].PID.UPD := 0.25, [0,11].PID.ERR := 0.20000005, [0,11].PID.MAXCV := 100.0, [0,11].PID.MAXTIE := 100.0, [0,11].PID.DATA[0] := -23.098158, [0,11].PID.DATA[3] := 0.20000005, [0,11].PID.DATA[4] := 0.20000005, [0,11].PID.DATA[5] := 0.024420025, [0,11].PID.DATA[6] := 1.0, [0,11].PID.DATA[7] := 4.0, [0,11].PID.DATA[8] := 0.1, [0,11].PID.DATA[9] := 0.1, [0,11].PID.DATA[11] := 0.1, [0,11].PID.DATA[12] := 0.1, [0,11].PID.DATA[15] := 1.0, [0,11].PID.DATA[16] := 1.0, [0,13].RampTimer.PRE := 3600000, [0,13].StableTimer.PRE := 2000, [0,13].PIDTimer.PRE := 10000, [0,13].PIDTimer.EN := 1, [0,13].PIDTimer.TT := 1, [0,13].PID.CTL := 305173120, [0,13].PID.PVT := 1, [0,13].PID.CA := 1, [0,13].PID.NOBC := 1, [0,13].PID.NOZC := 1, [0,13].PID.INI := 1, [0,13].PID.OLH := 1, [0,13].PID.DVPA := 1, [0,13].PID.PVHA := 1, [0,13].PID.KP := 0.2, [0,13].PID.KI := 0.08, [0,13].PID.MAXS := 100.0, [0,13].PID.DB := 1.0, [0,13].PID.SO := 100.0, [0,13].PID.MAXO := 100.0, [0,13].PID.UPD := 0.01, [0,13].PID.PV := 43.925232, [0,13].PID.ERR := 43.925232, [0,13].PID.OUT := 100.0, [0,13].PID.MAXI := 100.0, [0,13].PID.TIE := 2.4420025, [0,13].PID.MAXCV := 100.0, [0,13].PID.MAXTIE := 4095.0, [0,13].PID.DATA[0] := 100.0, [0,13].PID.DATA[1] := 702.8037, [0,13].PID.DATA[2] := 43.925232, [0,13].PID.DATA[3] := 43.925232, [0,13].PID.DATA[5] := 1.0, [0,13].PID.DATA[6] := 1.0, [0,13].PID.DATA[7] := 0.16, [0,13].PID.DATA[8] := 0.2, [0,13].PID.DATA[9] := 0.08, [0,13].PID.DATA[11] := 0.2, [0,13].PID.DATA[12] := 0.08,
        [0,13].PID.DATA[15] := 1.0, [0,13].PID.DATA[16] := 0.024420025, [1,0].RampTimer.PRE := 3600000, [1,0].StableTimer.PRE := 5000, [1,0].PIDTimer.PRE := 250, [1,0].PIDTimer.ACC := 100, [1,0].PIDTimer.EN := 1, [1,0].PIDTimer.TT := 1, [1,0].PID.CTL := 25199488, [1,0].PID.MO := 1, [1,0].PID.PE := 1, [1,0].PID.INI := 1, [1,0].PID.DVPA := 1, [1,0].PID.PVLA := 1, [1,0].PID.PVHA := 1, [1,0].PID.SP := 66.66666, [1,0].PID.KP := 0.5, [1,0].PID.KI := 0.1, [1,0].PID.MAXS := 200.0, [1,0].PID.SO := 10.0, [1,0].PID.MAXO := 100.0, [1,0].PID.MINO := 10.0, [1,0].PID.UPD := 0.25, [1,0].PID.ERR := 66.66666, [1,0].PID.OUT := 10.0, [1,0].PID.MAXI := 200.0, [1,0].PID.TIE := 10.0, [1,0].PID.MAXCV := 100.0, [1,0].PID.MAXTIE := 100.0, [1,0].PID.DATA[0] := -6.666666, [1,0].PID.DATA[3] := 66.66666, [1,0].PID.DATA[4] := 66.66666, [1,0].PID.DATA[5] := 0.5, [1,0].PID.DATA[6] := 1.0, [1,0].PID.DATA[7] := 4.0, [1,0].PID.DATA[8] := 0.5, [1,0].PID.DATA[9] := 0.1, [1,0].PID.DATA[11] := 0.5, [1,0].PID.DATA[12] := 0.08333334, [1,0].PID.DATA[15] := 1.0, [1,0].PID.DATA[16] := 1.0, [1,1].Tag := 'FIC01', [1,1].Desc := 'Feed Pump Control', [1,1].LoopCfg := 1, [1,1].ManualEGU := '%', [1,1].Manual := 1, [1,1].RampEnable := 1, [1,1].PIDEnable := 1, [1,1].ManualOSR := 1, [1,1].RangeMax := 100.0, [1,1].RampRate := 5.0, [1,1].RampRateSave := 5.0, [1,1].Deadband := 5.0, [1,1].RampTimer.PRE := 3600000, [1,1].StableTimer.PRE := 10000, [1,1].StableTime := 10, [1,1].PIDTimer.PRE := 250, [1,1].PIDTimer.EN := 1, [1,1].PIDTimer.TT := 1, [1,1].CycleTimer.PRE := 2000,
        [1,1].PID.CTL := 67143552, [1,1].PID.SWM := 1, [1,1].PID.INI := 1, [1,1].PID.DVNA := 1, [1,1].PID.DVPA := 1, [1,1].PID.PVLA := 1, [1,1].PID.PVHA := 1, [1,1].PID.KP := 0.1, [1,1].PID.KI := 0.2, [1,1].PID.MAXS := 25.0, [1,1].PID.DB := 0.01, [1,1].PID.MAXO := 100.0, [1,1].PID.UPD := 0.25, [1,1].PID.MAXI := 25.0, [1,1].PID.MAXCV := 100.0, [1,1].PID.MAXTIE := 25.0, [1,1].PID.DATA[5] := 4.0, [1,1].PID.DATA[6] := 1.0, [1,1].PID.DATA[7] := 4.0, [1,1].PID.DATA[8] := 0.1, [1,1].PID.DATA[9] := 0.2, [1,1].PID.DATA[11] := 0.1, [1,1].PID.DATA[12] := 0.2, [1,1].PID.DATA[15] := 1.0, [1,1].PID.DATA[16] := 4.0, [1,1].KP[0] := 100.0, [1,1].KP[1] := 100.0, [1,1].KI[0] := 200.0, [1,1].KI[1] := 200.0, [1,1].DB[0] := 0.01, [1,1].DB[1] := 0.01, [1,1].DB[2] := 0.01, [1,1].Auto1Cfg := 1, [1,1].Auto2Cfg := 1, [1,1].Auto1PVCfg := 42, [1,1].Auto2PVCfg := 40, [1,1].Auto1RangeMax := 25.0, [1,1].Auto2RangeMax := 6.0, [1,1].OutputAddress := 2, [1,2].Tag := 'LIC01', [1,2].Desc := 'Feed Bag Level', [1,2].LoopCfg := 1, [1,2].ManualEGU := '%', [1,2].Interlock := 1, [1,2].Manual := 1, [1,2].RampEnable := 1, [1,2].PIDEnable := 1, [1,2].ManualOSR := 1, [1,2].PVAuto1 := -0.16, [1,2].PVAuto2 := 2400.0, [1,2].RangeMax := 100.0, [1,2].RampRate := 5.0, [1,2].RampRateSave := 5.0, [1,2].Deadband := 5.0, [1,2].RampTimer.PRE := 3600000, [1,2].StableTimer.PRE := 10000, [1,2].StableTime := 10, [1,2].PIDTimer.PRE := 250, [1,2].PIDTimer.ACC := 95, [1,2].PIDTimer.EN := 1,
        [1,2].PIDTimer.TT := 1, [1,2].CycleTimer.PRE := 2000, [1,2].PID.CTL := 67143552, [1,2].PID.SWM := 1, [1,2].PID.INI := 1, [1,2].PID.DVNA := 1, [1,2].PID.DVPA := 1, [1,2].PID.PVLA := 1, [1,2].PID.PVHA := 1, [1,2].PID.KP := 5.0, [1,2].PID.KI := 10.0, [1,2].PID.MAXS := 50.0, [1,2].PID.DB := 0.001, [1,2].PID.MAXO := 100.0, [1,2].PID.UPD := 0.25, [1,2].PID.MAXI := 50.0, [1,2].PID.MAXCV := 100.0, [1,2].PID.MAXTIE := 100.0, [1,2].PID.DATA[5] := 2.0, [1,2].PID.DATA[6] := 1.0, [1,2].PID.DATA[7] := 4.0, [1,2].PID.DATA[8] := 5.0, [1,2].PID.DATA[9] := 10.0, [1,2].PID.DATA[11] := 5.0, [1,2].PID.DATA[12] := 10.0, [1,2].PID.DATA[15] := 1.0, [1,2].PID.DATA[16] := 1.0, [1,2].KP[0] := 5000.0, [1,2].KP[1] := 5000.0, [1,2].KI[0] := 10000.0, [1,2].KI[1] := 10000.0, [1,2].DB[0] := 0.001, [1,2].DB[1] := 0.001, [1,2].DB[2] := 0.001, [1,2].DisOSR := 1, [1,2].Auto1Cfg := 1, [1,2].Auto1PVCfg := 44, [1,2].Auto1RangeMax := 50.0, [1,2].OutputAddress := 3, [1,3].Tag := 'PCV01', [1,3].Desc := 'Retentate control valve', [1,3].LoopCfg := 1, [1,3].ManualEGU := '%', [1,3].Enable := 1, [1,3].Manual := 1, [1,3].Stable := 1, [1,3].Status := 1, [1,3].RampEnable := 1, [1,3].PIDEnable := 1, [1,3].ManualOSR := 1, [1,3].PV := -0.03822385, [1,3].PVAuto1 := -0.03822385, [1,3].SPAutoSave := -0.03822385, [1,3].RangeMax := 100.0, [1,3].RampRate := 5.0, [1,3].RampRateSave := 5.0, [1,3].Deadband := 10.0, [1,3].RampTimer.PRE := 3600000, [1,3].StableTimer.PRE := 5000, [1,3].StableTime := 5,
        [1,3].PIDTimer.PRE := 250, [1,3].PIDTimer.EN := 1, [1,3].PIDTimer.TT := 1, [1,3].CycleTimer.PRE := 2000, [1,3].PID.CTL := 67142400, [1,3].PID.SWM := 1, [1,3].PID.INI := 1, [1,3].PID.DVPA := 1, [1,3].PID.PVLA := 1, [1,3].PID.KP := 0.04, [1,3].PID.KI := 0.04, [1,3].PID.BIAS := 30.796, [1,3].PID.MAXS := 6.0, [1,3].PID.DB := 0.02, [1,3].PID.MAXO := 100.0, [1,3].PID.UPD := 0.25, [1,3].PID.PV := -0.03730831, [1,3].PID.ERR := 0.03730831, [1,3].PID.MAXI := 6.0, [1,3].PID.MAXCV := 100.0, [1,3].PID.MAXTIE := 100.0, [1,3].PID.DATA[0] := -30.820871, [1,3].PID.DATA[1] := 9.948882, [1,3].PID.DATA[2] := -0.03730831, [1,3].PID.DATA[3] := 0.03730831, [1,3].PID.DATA[5] := 16.666666, [1,3].PID.DATA[6] := 1.0, [1,3].PID.DATA[7] := 4.0, [1,3].PID.DATA[8] := 0.04, [1,3].PID.DATA[9] := 0.04, [1,3].PID.DATA[11] := 0.04, [1,3].PID.DATA[12] := 0.04, [1,3].PID.DATA[15] := 1.0, [1,3].PID.DATA[16] := 1.0, [1,3].KP[0] := 40.0, [1,3].KP[1] := 40.0, [1,3].KI[0] := 40.0, [1,3].KI[1] := 40.0, [1,3].DB[0] := 0.02, [1,3].DB[1] := 0.02, [1,3].Auto1Cfg := 1, [1,3].Auto2Cfg := 1, [1,3].Auto1PVCfg := 6, [1,3].Auto2PVCfg := 41, [1,3].Auto1RangeMax := 6.0, [1,3].Auto2RangeMax := 6.0, [1,4].ManualEGU := '%', [1,4].Enable := 1, [1,4].Status := 3, [1,4].PIDEnable := 1, [1,4].PV := 101.99314, [1,4].PVAuto1 := -1.4998856, [1,4].SPAutoSave := -1.4998856, [1,4].RangeMax := 100.0, [1,4].RampRate := 6.0, [1,4].RampRateSave := 6.0, [1,4].Deadband := 2.0, [1,4].RampTimer.PRE := 3600000, [1,4].StableTimer.PRE := 10000, [1,4].StableTime := 5,
        [1,4].PIDTimer.PRE := 250, [1,4].CycleTimer.PRE := 2000, [1,4].PID.CTL := -2145344384, [1,4].PID.EN := 1, [1,4].PID.NOBC := 1, [1,4].PID.INI := 1, [1,4].PID.OLL := 1, [1,4].PID.DVNA := 1, [1,4].PID.PVHA := 1, [1,4].PID.KP := 0.2, [1,4].PID.KI := 0.08, [1,4].PID.KD := 0.01, [1,4].PID.MAXS := 100.0, [1,4].PID.DB := 0.3, [1,4].PID.MAXO := 100.0, [1,4].PID.UPD := 0.005, [1,4].PID.PV := 101.99314, [1,4].PID.ERR := -101.99314, [1,4].PID.MAXI := 100.0, [1,4].PID.MAXCV := 100.0, [1,4].PID.MAXTIE := 4095.0, [1,4].PID.DATA[0] := -105.9066, [1,4].PID.DATA[1] := -1631.9136, [1,4].PID.DATA[2] := 101.99314, [1,4].PID.DATA[3] := -101.99314, [1,4].PID.DATA[5] := 1.0, [1,4].PID.DATA[6] := 1.0, [1,4].PID.DATA[7] := 0.089999996, [1,4].PID.DATA[8] := 0.2, [1,4].PID.DATA[9] := 0.08, [1,4].PID.DATA[10] := 0.01, [1,4].PID.DATA[11] := 0.2, [1,4].PID.DATA[12] := 0.08, [1,4].PID.DATA[13] := 0.01, [1,4].PID.DATA[15] := 1.0, [1,4].PID.DATA[16] := 0.024420025, [1,5].Tag := 'PCV11', [1,5].Desc := 'Filtrate control valve', [1,5].LoopCfg := 1, [1,5].ManualEGU := '%', [1,5].Enable := 1, [1,5].Manual := 1, [1,5].Stable := 1, [1,5].Status := 2, [1,5].RampEnable := 1, [1,5].PIDEnable := 1, [1,5].ManualOSR := 1, [1,5].PV := 0.01201648, [1,5].PVAuto1 := 0.01201648, [1,5].SPAutoSave := 0.01201648, [1,5].RangeMax := 100.0, [1,5].RampRate := 5.0, [1,5].RampRateSave := 5.0, [1,5].RampStart := 4.417, [1,5].Deadband := 10.0, [1,5].RampTimer.PRE := 3600000, [1,5].StableTimer.PRE := 5000, [1,5].StableTime := 5, [1,5].PIDTimer.PRE := 250, [1,5].PIDTimer.ACC := 188,
        [1,5].PIDTimer.EN := 1, [1,5].PIDTimer.TT := 1, [1,5].CycleTimer.PRE := 2000, [1,5].PID.CTL := 67142784, [1,5].PID.SWM := 1, [1,5].PID.INI := 1, [1,5].PID.DVNA := 1, [1,5].PID.PVHA := 1, [1,5].PID.KP := 0.25, [1,5].PID.KI := 0.01, [1,5].PID.KD := 0.01, [1,5].PID.BIAS := -847.4798, [1,5].PID.MAXS := 15.0, [1,5].PID.DB := 0.02, [1,5].PID.MAXO := 100.0, [1,5].PID.UPD := 0.25, [1,5].PID.PV := 0.014305333, [1,5].PID.ERR := -0.014305333, [1,5].PID.MAXI := 15.0, [1,5].PID.MAXCV := 100.0, [1,5].PID.MAXTIE := 100.0, [1,5].PID.DATA[0] := 847.5043, [1,5].PID.DATA[1] := -1.5252948, [1,5].PID.DATA[2] := 0.014305333, [1,5].PID.DATA[3] := -0.014305333, [1,5].PID.DATA[5] := 6.6666665, [1,5].PID.DATA[6] := 1.0, [1,5].PID.DATA[7] := 4.01, [1,5].PID.DATA[8] := 0.25, [1,5].PID.DATA[9] := 0.01, [1,5].PID.DATA[10] := 0.01, [1,5].PID.DATA[11] := 0.25, [1,5].PID.DATA[12] := 0.01, [1,5].PID.DATA[13] := 0.01, [1,5].PID.DATA[15] := 1.0, [1,5].PID.DATA[16] := 1.0, [1,5].KP[0] := 250.0, [1,5].KP[1] := 250.0, [1,5].KI[0] := 10.0, [1,5].KI[1] := 10.0, [1,5].KD[0] := 10.0, [1,5].KD[1] := 10.0, [1,5].DB[0] := 0.02, [1,5].DB[1] := 0.02, [1,5].Auto1Cfg := 1, [1,5].Auto2Cfg := 1, [1,5].Auto1PVCfg := 2, [1,5].Auto2PVCfg := 41, [1,5].Auto1RangeMax := 15.0, [1,5].Auto2RangeMax := 6.0, [1,5].OutputAddress := 1, [1,6].Enable := 1, [1,6].Stable := 1, [1,6].Status := 3, [1,6].PIDEnable := 1, [1,6].PV := 38.696636, [1,6].PVAuto1 := -3.749714, [1,6].PVAuto2 := 1.9581139, [1,6].SPAutoSave := -3.749714, [1,6].RangeMax := 100.0,
        [1,6].RampRate := 6.0, [1,6].RampRateSave := 6.0, [1,6].Deadband := 2.0, [1,6].RampTimer.PRE := 3600000, [1,6].StableTimer.PRE := 5000, [1,6].StableTime := 5, [1,6].PIDTimer.PRE := 250, [1,6].CycleTimer.PRE := 2000, [1,6].PID.CTL := -2145344384, [1,6].PID.EN := 1, [1,6].PID.NOBC := 1, [1,6].PID.INI := 1, [1,6].PID.OLL := 1, [1,6].PID.DVNA := 1, [1,6].PID.PVHA := 1, [1,6].PID.KP := 0.3, [1,6].PID.KI := 0.25, [1,6].PID.KD := 0.01, [1,6].PID.MAXS := 100.0, [1,6].PID.DB := 0.3, [1,6].PID.MAXO := 100.0, [1,6].PID.UPD := 0.005, [1,6].PID.PV := 38.696636, [1,6].PID.ERR := -38.696636, [1,6].PID.MAXI := 100.0, [1,6].PID.MAXCV := 100.0, [1,6].PID.MAXTIE := 4095.0, [1,6].PID.DATA[0] := 11.461082, [1,6].PID.DATA[1] := -619.0884, [1,6].PID.DATA[2] := 38.696636, [1,6].PID.DATA[3] := -38.696636, [1,6].PID.DATA[5] := 1.0, [1,6].PID.DATA[6] := 1.0, [1,6].PID.DATA[7] := 0.089999996, [1,6].PID.DATA[8] := 0.3, [1,6].PID.DATA[9] := 0.25, [1,6].PID.DATA[10] := 0.01, [1,6].PID.DATA[11] := 0.3, [1,6].PID.DATA[12] := 0.25, [1,6].PID.DATA[13] := 0.01, [1,6].PID.DATA[15] := 1.0, [1,6].PID.DATA[16] := 0.024420025, [1,6].OutputAddress := 1, [1,7].StableTimer.PRE := 200, [1,7].PIDTimer.PRE := 250, [1,7].PIDTimer.EN := 1, [1,7].PIDTimer.TT := 1, [1,7].CycleTimer.PRE := 10000, [1,7].PID.CTL := 16810880, [1,7].PID.MO := 1, [1,7].PID.INI := 1, [1,7].PID.DVPA := 1, [1,7].PID.PVLA := 1, [1,7].PID.PVHA := 1, [1,7].PID.SP := 10.0, [1,7].PID.KP := 2.0, [1,7].PID.KI := 0.2, [1,7].PID.KD := 0.3, [1,7].PID.BIAS := 50.0, [1,7].PID.DB := 0.01,
        [1,7].PID.SO := 80.0, [1,7].PID.MAXO := 100.0, [1,7].PID.UPD := 0.25, [1,7].PID.ERR := 10.0, [1,7].PID.OUT := 80.0, [1,7].PID.TIE := 80.0, [1,7].PID.MAXCV := 100.0, [1,7].PID.MAXTIE := 100.0, [1,7].PID.DATA[0] := 29.511597, [1,7].PID.DATA[3] := 10.0, [1,7].PID.DATA[4] := 10.0, [1,7].PID.DATA[5] := 0.024420025, [1,7].PID.DATA[6] := 1.0, [1,7].PID.DATA[7] := 4.3, [1,7].PID.DATA[8] := 2.0, [1,7].PID.DATA[9] := 0.2, [1,7].PID.DATA[10] := 0.3, [1,7].PID.DATA[11] := 2.0, [1,7].PID.DATA[12] := 0.2, [1,7].PID.DATA[13] := 0.3, [1,7].PID.DATA[15] := 1.0, [1,7].PID.DATA[16] := 1.0, [1,8].StableTimer.PRE := 15000, [1,8].PIDTimer.PRE := 250, [1,8].CycleTimer.PRE := 20000, [1,8].PID.CTL := 33555584, [1,8].PID.CA := 1, [1,8].PID.DVNA := 1, [1,8].PID.PVHA := 1, [1,8].PID.SP := 27.0, [1,8].PID.KP := 1.0, [1,8].PID.KI := 0.1, [1,8].PID.MAXS := 100.0, [1,8].PID.MAXO := 100.0, [1,8].PID.UPD := 0.25, [1,8].PID.PV := 18.2328, [1,8].PID.ERR := -8.767202, [1,8].PID.MAXI := 100.0, [1,8].PID.MAXCV := 100.0, [1,8].PID.MAXTIE := 100.0, [1,8].PID.DATA[0] := 8.767202, [1,8].PID.DATA[1] := 291.7248, [1,8].PID.DATA[2] := 18.2328, [1,8].PID.DATA[3] := -8.767202, [1,8].PID.DATA[4] := 27.0, [1,8].PID.DATA[5] := 1.0, [1,8].PID.DATA[6] := 1.0, [1,8].PID.DATA[7] := 4.0, [1,8].PID.DATA[8] := 1.0, [1,8].PID.DATA[9] := 0.1, [1,8].PID.DATA[11] := 1.0, [1,8].PID.DATA[12] := 0.1, [1,8].PID.DATA[15] := 1.0, [1,8].PID.DATA[16] := 1.0, [1,11].RampTimer.PRE := 100000, [1,11].StableTimer.PRE := 200, [1,11].PIDTimer.PRE := 250, [1,11].PIDTimer.ACC := 230, [1,11].PIDTimer.EN := 1, [1,11].PIDTimer.TT := 1,
        [1,11].PID.CTL := 67142528, [1,11].PID.SWM := 1, [1,11].PID.INI := 1, [1,11].PID.DVPA := 1, [1,11].PID.PVLA := 1, [1,11].PID.PVHA := 1, [1,11].PID.SP := 0.20000005, [1,11].PID.KP := 0.1, [1,11].PID.KI := 0.1, [1,11].PID.BIAS := 23.09767, [1,11].PID.DB := 0.001, [1,11].PID.MAXO := 100.0, [1,11].PID.UPD := 0.25, [1,11].PID.ERR := 0.20000005, [1,11].PID.MAXCV := 100.0, [1,11].PID.MAXTIE := 100.0, [1,11].PID.DATA[0] := -23.098158, [1,11].PID.DATA[3] := 0.20000005, [1,11].PID.DATA[4] := 0.20000005, [1,11].PID.DATA[5] := 0.024420025, [1,11].PID.DATA[6] := 1.0, [1,11].PID.DATA[7] := 4.0, [1,11].PID.DATA[8] := 0.1, [1,11].PID.DATA[9] := 0.1, [1,11].PID.DATA[11] := 0.1, [1,11].PID.DATA[12] := 0.1, [1,11].PID.DATA[15] := 1.0, [1,11].PID.DATA[16] := 1.0, [1,12].Enable := 1, [1,12].Manual := 1, [1,12].Stable := 1, [1,12].RampEnable := 1, [1,12].PIDEnable := 1, [1,12].ManualOSR := 1, [1,12].PV := 54.98666, [1,12].SPAutoSave := 54.98666, [1,12].SPManual := 50.0, [1,12].SPManualSave := 50.0, [1,12].RampRate := 0.5, [1,12].RampRateSave := 0.5, [1,12].RampStart := 34.736, [1,12].Deadband := 6.6, [1,12].RampTimer.PRE := 3600000, [1,12].PIDTimer.EN := 1, [1,12].PIDTimer.TT := 1, [1,12].PID.CTL := 67141632, [1,12].PID.SWM := 1, [1,12].PID.INI := 1, [1,12].PID.KP := 0.2, [1,12].PID.KI := 0.2, [1,12].PID.MAXS := 50.0, [1,12].PID.SO := 6.4153447, [1,12].PID.MAXO := 100.0, [1,12].PID.MAXI := 50.0, [1,12].PID.MAXTIE := 4095.0, [1,12].PID.DATA[5] := 2.0, [1,12].PID.DATA[6] := 1.0, [1,12].PID.DATA[16] := 0.024420025, [1,12].DisOSR := 1, [1,12].Auto1Cfg := 1,
        [1,12].Auto2Cfg := 1, [1,12].Auto1PVCfg := 1, [1,12].Auto2PVCfg := 33, [1,12].Auto3PVCfg := 1, [1,12].OutputAddress := 2, [1,13].Enable := 1, [1,13].Stable := 1, [1,13].DBOK := 1, [1,13].PIDEnable := 1, [1,13].PV := 100.545425, [1,13].CV := 6.5049314, [1,13].SPAuto := 100.0, [1,13].RampRate := 0.6, [1,13].RampRateSave := 0.6, [1,13].RampStart := 100.0, [1,13].Deadband := 2.0, [1,13].DBLO := 98.0, [1,13].DBHI := 102.0, [1,13].RampTimer.PRE := 3600000, [1,13].StableTimer.PRE := 2000, [1,13].StableTimer.ACC := 2000, [1,13].StableTimer.EN := 1, [1,13].StableTimer.DN := 1, [1,13].PIDTimer.PRE := 10000, [1,13].PID.CTL := -2111798656, [1,13].PID.EN := 1, [1,13].PID.CA := 1, [1,13].PID.NOBC := 1, [1,13].PID.INI := 1, [1,13].PID.DVPA := 1, [1,13].PID.PVHA := 1, [1,13].PID.SP := 100.0, [1,13].PID.KP := 0.2, [1,13].PID.KI := 0.25, [1,13].PID.KD := 0.01, [1,13].PID.MAXS := 100.0, [1,13].PID.DB := 0.3, [1,13].PID.SO := 6.5049314, [1,13].PID.MAXO := 100.0, [1,13].PID.UPD := 0.005, [1,13].PID.PV := 100.545425, [1,13].PID.ERR := 0.5454254, [1,13].PID.OUT := 6.5049314, [1,13].PID.MAXI := 100.0, [1,13].PID.TIE := 0.15657456, [1,13].PID.MAXCV := 100.0, [1,13].PID.MAXTIE := 4095.0, [1,13].PID.DATA[0] := 6.3127437, [1,13].PID.DATA[1] := 1608.6437, [1,13].PID.DATA[2] := 100.545425, [1,13].PID.DATA[3] := 0.5454254, [1,13].PID.DATA[4] := 100.0, [1,13].PID.DATA[5] := 1.0, [1,13].PID.DATA[6] := 1.0, [1,13].PID.DATA[7] := 0.089999996, [1,13].PID.DATA[8] := 0.2, [1,13].PID.DATA[9] := 0.25, [1,13].PID.DATA[10] := 0.01, [1,13].PID.DATA[11] := 0.2, [1,13].PID.DATA[12] := 0.25,
        [1,13].PID.DATA[13] := 0.01, [1,13].PID.DATA[15] := 1.0, [1,13].PID.DATA[16] := 0.024420025, [1,13].OutputAddress := 2, [2,0].RampTimer.PRE := 3600000, [2,0].StableTimer.PRE := 5000, [2,0].PIDTimer.PRE := 250, [2,0].PIDTimer.ACC := 100, [2,0].PIDTimer.EN := 1, [2,0].PIDTimer.TT := 1, [2,0].PID.CTL := 25199488, [2,0].PID.MO := 1, [2,0].PID.PE := 1, [2,0].PID.INI := 1, [2,0].PID.DVPA := 1, [2,0].PID.PVLA := 1, [2,0].PID.PVHA := 1, [2,0].PID.SP := 66.66666, [2,0].PID.KP := 0.5, [2,0].PID.KI := 0.1, [2,0].PID.MAXS := 200.0, [2,0].PID.SO := 10.0, [2,0].PID.MAXO := 100.0, [2,0].PID.MINO := 10.0, [2,0].PID.UPD := 0.25, [2,0].PID.ERR := 66.66666, [2,0].PID.OUT := 10.0, [2,0].PID.MAXI := 200.0, [2,0].PID.TIE := 10.0, [2,0].PID.MAXCV := 100.0, [2,0].PID.MAXTIE := 100.0, [2,0].PID.DATA[0] := -6.666666, [2,0].PID.DATA[3] := 66.66666, [2,0].PID.DATA[4] := 66.66666, [2,0].PID.DATA[5] := 0.5, [2,0].PID.DATA[6] := 1.0, [2,0].PID.DATA[7] := 4.0, [2,0].PID.DATA[8] := 0.5, [2,0].PID.DATA[9] := 0.1, [2,0].PID.DATA[11] := 0.5, [2,0].PID.DATA[12] := 0.08333334, [2,0].PID.DATA[15] := 1.0, [2,0].PID.DATA[16] := 1.0, [2,1].Tag := 'FIC01', [2,1].Desc := 'Feed Pump Control Loop', [2,1].LoopCfg := 1, [2,1].ManualEGU := '%', [2,1].Auto1EGU := 'LPM', [2,1].Auto2EGU := 'Bar', [2,1].Manual := 1, [2,1].DBOK := 1, [2,1].RampEnable := 1, [2,1].PIDEnable := 1, [2,1].ManualOSR := 1, [2,1].PVAuto2 := 2400.0, [2,1].RangeMax := 100.0, [2,1].RampRate := 5.0, [2,1].RampRateSave := 5.0, [2,1].Deadband := 5.0, [2,1].RampTimer.PRE := 3600000,
        [2,1].StableTimer.PRE := 10000, [2,1].StableTime := 10, [2,1].PIDTimer.PRE := 250, [2,1].PIDTimer.EN := 1, [2,1].PIDTimer.TT := 1, [2,1].CycleTimer.PRE := 2000, [2,1].PID.CTL := 67143552, [2,1].PID.SWM := 1, [2,1].PID.INI := 1, [2,1].PID.DVNA := 1, [2,1].PID.DVPA := 1, [2,1].PID.PVLA := 1, [2,1].PID.PVHA := 1, [2,1].PID.KP := 0.1, [2,1].PID.KI := 0.2, [2,1].PID.MAXS := 45.0, [2,1].PID.DB := 0.01, [2,1].PID.MAXO := 100.0, [2,1].PID.UPD := 0.25, [2,1].PID.MAXI := 45.0, [2,1].PID.MAXCV := 100.0, [2,1].PID.MAXTIE := 45.0, [2,1].PID.DATA[5] := 2.2222223, [2,1].PID.DATA[6] := 1.0, [2,1].PID.DATA[7] := 4.0, [2,1].PID.DATA[8] := 0.1, [2,1].PID.DATA[9] := 0.2, [2,1].PID.DATA[11] := 0.1, [2,1].PID.DATA[12] := 0.2, [2,1].PID.DATA[15] := 1.0, [2,1].PID.DATA[16] := 2.2222223, [2,1].KP[0] := 100.0, [2,1].KP[1] := 100.0, [2,1].KI[0] := 200.0, [2,1].KI[1] := 200.0, [2,1].DB[0] := 0.01, [2,1].Auto1Cfg := 1, [2,1].Auto2Cfg := 1, [2,1].Auto1PVCfg := 42, [2,1].Auto2PVCfg := 40, [2,1].Auto1RangeMax := 45.0, [2,1].Auto2RangeMax := 6.0, [2,1].OutputAddress := 2, [2,2].Tag := 'LIC01', [2,2].Desc := 'Level Control Loop', [2,2].LoopCfg := 1, [2,2].ManualEGU := '%', [2,2].Auto1EGU := 'L', [2,2].Interlock := 1, [2,2].Manual := 1, [2,2].DBOK := 1, [2,2].RampEnable := 1, [2,2].PIDEnable := 1, [2,2].ManualOSR := 1, [2,2].PVAuto2 := 2400.0, [2,2].RangeMax := 100.0, [2,2].RampRate := 5.0, [2,2].RampRateSave := 5.0, [2,2].RampStart := 75.0, [2,2].Deadband := 5.0,
        [2,2].RampTimer.PRE := 3600000, [2,2].StableTimer.PRE := 10000, [2,2].StableTime := 10, [2,2].PIDTimer.PRE := 250, [2,2].PIDTimer.EN := 1, [2,2].PIDTimer.TT := 1, [2,2].CycleTimer.PRE := 2000, [2,2].PID.CTL := 67143552, [2,2].PID.SWM := 1, [2,2].PID.INI := 1, [2,2].PID.DVNA := 1, [2,2].PID.DVPA := 1, [2,2].PID.PVLA := 1, [2,2].PID.PVHA := 1, [2,2].PID.KP := 5.0, [2,2].PID.KI := 10.0, [2,2].PID.MAXS := 50.0, [2,2].PID.DB := 0.001, [2,2].PID.MAXO := 100.0, [2,2].PID.UPD := 0.25, [2,2].PID.MAXI := 50.0, [2,2].PID.MAXCV := 100.0, [2,2].PID.MAXTIE := 100.0, [2,2].PID.DATA[5] := 2.0, [2,2].PID.DATA[6] := 1.0, [2,2].PID.DATA[7] := 4.0, [2,2].PID.DATA[8] := 5.0, [2,2].PID.DATA[9] := 10.0, [2,2].PID.DATA[11] := 5.0, [2,2].PID.DATA[12] := 10.0, [2,2].PID.DATA[15] := 1.0, [2,2].PID.DATA[16] := 1.0, [2,2].KP[0] := 5000.0, [2,2].KP[1] := 5000.0, [2,2].KI[0] := 10000.0, [2,2].KI[1] := 10000.0, [2,2].DB[0] := 0.001, [2,2].DisOSR := 1, [2,2].Auto1Cfg := 1, [2,2].Auto1PVCfg := 44, [2,2].Auto1RangeMax := 50.0, [2,2].OutputAddress := 3, [2,3].Tag := 'Mixer', [2,3].ManualEGU := '%', [2,3].Enable := 1, [2,3].Manual := 1, [2,3].Stable := 1, [2,3].DBOK := 1, [2,3].Status := 3, [2,3].RampEnable := 1, [2,3].PIDEnable := 1, [2,3].ManualOSR := 1, [2,3].RangeMax := 100.0, [2,3].RampRate := 5.0, [2,3].RampRateSave := 5.0, [2,3].RampStart := 98.0, [2,3].Deadband := 10.0, [2,3].RampTimer.PRE := 3600000, [2,3].StableTimer.PRE := 2300, [2,3].StableTimer.ACC := 2354,
        [2,3].StableTimer.EN := 1, [2,3].StableTimer.DN := 1, [2,3].StableTime := 10, [2,3].PIDTimer.PRE := 250, [2,3].PIDTimer.ACC := 214, [2,3].PIDTimer.EN := 1, [2,3].PIDTimer.TT := 1, [2,3].CycleTimer.PRE := 2000, [2,3].PID.CTL := 67110784, [2,3].PID.SWM := 1, [2,3].PID.DVNA := 1, [2,3].PID.DVPA := 1, [2,3].PID.PVLA := 1, [2,3].PID.PVHA := 1, [2,3].PID.KP := 0.001, [2,3].PID.KI := 0.001, [2,3].PID.BIAS := 30.796, [2,3].PID.MAXS := 4095.0, [2,3].PID.DB := 0.02, [2,3].PID.MAXO := 100.0, [2,3].PID.UPD := 0.25, [2,3].PID.MAXI := 4095.0, [2,3].PID.MAXCV := 100.0, [2,3].PID.MAXTIE := 100.0, [2,3].PID.DATA[0] := -30.796, [2,3].PID.DATA[5] := 0.024420025, [2,3].PID.DATA[6] := 1.0, [2,3].PID.DATA[7] := 0.16, [2,3].PID.DATA[8] := 0.001, [2,3].PID.DATA[9] := 0.001, [2,3].PID.DATA[11] := 0.001, [2,3].PID.DATA[12] := 0.001, [2,3].PID.DATA[15] := 1.0, [2,3].PID.DATA[16] := 1.0, [2,3].KP[0] := 40.0, [2,3].KP[1] := 40.0, [2,3].KI[0] := 40.0, [2,3].KI[1] := 40.0, [2,3].DB[0] := 0.02, [2,3].DB[1] := 0.02, [2,3].OutputAddress := 2, [2,4].Tag := 'PC001', [2,4].Desc := 'Retentate Control Valve', [2,4].LoopCfg := 1, [2,4].ManualEGU := '%', [2,4].Auto1EGU := 'Bar', [2,4].Auto2EGU := 'Bar', [2,4].Enable := 1, [2,4].Manual := 1, [2,4].Stable := 1, [2,4].Status := 3, [2,4].RampEnable := 1, [2,4].PIDEnable := 1, [2,4].ManualOSR := 1, [2,4].PV := -1.4998856, [2,4].PVAuto1 := -1.4998856, [2,4].SPAutoSave := -1.4998856, [2,4].RangeMax := 100.0, [2,4].RampRate := 1.0, [2,4].RampRateSave := 1.0,
        [2,4].Deadband := 10.0, [2,4].RampTimer.PRE := 3600000, [2,4].StableTimer.PRE := 5000, [2,4].StableTime := 5, [2,4].PIDTimer.PRE := 250, [2,4].CycleTimer.PRE := 2000, [2,4].PID.CTL := -2078276864, [2,4].PID.EN := 1, [2,4].PID.SWM := 1, [2,4].PID.NOBC := 1, [2,4].PID.DVPA := 1, [2,4].PID.PVLA := 1, [2,4].PID.KP := 0.04, [2,4].PID.KI := 0.001, [2,4].PID.KD := 0.02, [2,4].PID.MAXS := 6.0, [2,4].PID.DB := 0.3, [2,4].PID.MAXO := 100.0, [2,4].PID.UPD := 0.25, [2,4].PID.PV := -1.4998856, [2,4].PID.ERR := 1.4998856, [2,4].PID.MAXI := 6.0, [2,4].PID.MAXCV := 100.0, [2,4].PID.MAXTIE := 4095.0, [2,4].PID.DATA[0] := -0.9999237, [2,4].PID.DATA[1] := 399.96948, [2,4].PID.DATA[2] := -1.4998856, [2,4].PID.DATA[3] := 1.4998856, [2,4].PID.DATA[5] := 16.666666, [2,4].PID.DATA[6] := 1.0, [2,4].PID.DATA[7] := 4.02, [2,4].PID.DATA[8] := 0.04, [2,4].PID.DATA[9] := 0.001, [2,4].PID.DATA[10] := 0.02, [2,4].PID.DATA[11] := 0.04, [2,4].PID.DATA[12] := 0.001, [2,4].PID.DATA[13] := 0.02, [2,4].PID.DATA[15] := 1.0, [2,4].PID.DATA[16] := 16.666666, [2,4].KP[0] := 40.0, [2,4].KP[1] := 40.0, [2,4].KI[0] := 1.0, [2,4].KI[1] := 40.0, [2,4].DB[0] := 0.02, [2,4].Auto1Cfg := 1, [2,4].Auto2Cfg := 1, [2,4].Auto1PVCfg := 6, [2,4].Auto2PVCfg := 41, [2,4].Auto1RangeMax := 6.0, [2,4].Auto2RangeMax := 6.0, [2,5].ManualEGU := '%', [2,5].Manual := 1, [2,5].Status := 3, [2,5].RampEnable := 1, [2,5].PIDEnable := 1, [2,5].RangeMax := 100.0, [2,5].RampRate := 5.0, [2,5].RampRateSave := 5.0, [2,5].RampStart := 4.417, [2,5].Deadband := 10.0,
        [2,5].RampTimer.PRE := 3600000, [2,5].StableTimer.PRE := 1500, [2,5].StableTime := 10, [2,5].PIDTimer.PRE := 250, [2,5].CycleTimer.PRE := 2000, [2,5].PID.CTL := 896, [2,5].PID.DVPA := 1, [2,5].PID.PVLA := 1, [2,5].PID.PVHA := 1, [2,5].PID.SP := 350.0, [2,5].PID.KP := 40.0, [2,5].PID.KI := 0.5, [2,5].PID.BIAS := -847.4798, [2,5].PID.MAXS := 550.0, [2,5].PID.MAXO := 100.0, [2,5].PID.UPD := 0.25, [2,5].PID.ERR := 350.0, [2,5].PID.MAXI := 550.0, [2,5].PID.MAXCV := 100.0, [2,5].PID.MAXTIE := 100.0, [2,5].PID.DATA[0] := -1697.975, [2,5].PID.DATA[1] := 1018.182, [2,5].PID.DATA[3] := 350.0, [2,5].PID.DATA[4] := 350.0, [2,5].PID.DATA[5] := 0.1818182, [2,5].PID.DATA[6] := 1.0, [2,5].PID.DATA[7] := 4.0, [2,5].PID.DATA[8] := 40.0, [2,5].PID.DATA[9] := 0.5, [2,5].PID.DATA[11] := 40.0, [2,5].PID.DATA[12] := 0.5, [2,5].PID.DATA[15] := 1.0, [2,5].PID.DATA[16] := 1.0, [2,5].KP[0] := 250.0, [2,5].KP[1] := 250.0, [2,5].KI[0] := 100.0, [2,5].KI[1] := 100.0, [2,5].KD[0] := 100.0, [2,5].KD[1] := 100.0, [2,5].DB[0] := 0.02, [2,5].DB[1] := 0.02, [2,5].OutputAddress := 3, [2,6].Tag := 'PC101', [2,6].Desc := 'Filtrate Control Valve', [2,6].LoopCfg := 1, [2,6].AutoEGU := 'Bar', [2,6].Auto1EGU := 'Bar', [2,6].Enable := 1, [2,6].Manual := 1, [2,6].Stable := 1, [2,6].Status := 3, [2,6].RampEnable := 1, [2,6].PIDEnable := 1, [2,6].ManualOSR := 1, [2,6].PV := -6.249523, [2,6].PVAuto1 := -6.249523, [2,6].SPAutoSave := -6.249523, [2,6].RangeMax := 100.0, [2,6].RampRate := 1.0, [2,6].RampRateSave := 1.0,
        [2,6].Deadband := 10.0, [2,6].RampTimer.PRE := 3600000, [2,6].StableTimer.PRE := 5000, [2,6].StableTime := 5, [2,6].PIDTimer.PRE := 250, [2,6].CycleTimer.PRE := 2000, [2,6].PID.CTL := -2078276864, [2,6].PID.EN := 1, [2,6].PID.SWM := 1, [2,6].PID.NOBC := 1, [2,6].PID.DVPA := 1, [2,6].PID.PVLA := 1, [2,6].PID.KP := 0.1, [2,6].PID.KI := 0.005, [2,6].PID.KD := 0.02, [2,6].PID.MAXS := 25.0, [2,6].PID.DB := 0.3, [2,6].PID.MAXO := 100.0, [2,6].PID.UPD := 0.25, [2,6].PID.PV := -6.249523, [2,6].PID.ERR := 6.249523, [2,6].PID.MAXI := 25.0, [2,6].PID.MAXCV := 100.0, [2,6].PID.MAXTIE := 4095.0, [2,6].PID.DATA[0] := -2.4998093, [2,6].PID.DATA[1] := 399.96948, [2,6].PID.DATA[2] := -6.249523, [2,6].PID.DATA[3] := 6.249523, [2,6].PID.DATA[5] := 4.0, [2,6].PID.DATA[6] := 1.0, [2,6].PID.DATA[7] := 4.02, [2,6].PID.DATA[8] := 0.1, [2,6].PID.DATA[9] := 0.005, [2,6].PID.DATA[10] := 0.02, [2,6].PID.DATA[11] := 0.1, [2,6].PID.DATA[12] := 0.005, [2,6].PID.DATA[13] := 0.02, [2,6].PID.DATA[15] := 1.0, [2,6].PID.DATA[16] := 4.0, [2,6].KP[0] := 100.0, [2,6].KP[1] := 250.0, [2,6].KI[0] := 5.0, [2,6].KI[1] := 20.0, [2,6].DB[0] := 0.02, [2,6].Auto1Cfg := 1, [2,6].Auto2Cfg := 1, [2,6].Auto1PVCfg := 2, [2,6].Auto2PVCfg := 41, [2,6].Auto1RangeMax := 25.0, [2,6].Auto2RangeMax := 6.0, [2,6].OutputAddress := 1, [2,7].StableTimer.PRE := 200, [2,7].PIDTimer.PRE := 250, [2,7].PIDTimer.EN := 1, [2,7].PIDTimer.TT := 1, [2,7].CycleTimer.PRE := 10000, [2,7].PID.CTL := 16810880, [2,7].PID.MO := 1, [2,7].PID.INI := 1, [2,7].PID.DVPA := 1,
        [2,7].PID.PVLA := 1, [2,7].PID.PVHA := 1, [2,7].PID.SP := 10.0, [2,7].PID.KP := 2.0, [2,7].PID.KI := 0.2, [2,7].PID.KD := 0.3, [2,7].PID.BIAS := 50.0, [2,7].PID.DB := 0.01, [2,7].PID.SO := 80.0, [2,7].PID.MAXO := 100.0, [2,7].PID.UPD := 0.25, [2,7].PID.ERR := 10.0, [2,7].PID.OUT := 80.0, [2,7].PID.TIE := 80.0, [2,7].PID.MAXCV := 100.0, [2,7].PID.MAXTIE := 100.0, [2,7].PID.DATA[0] := 29.5116, [2,7].PID.DATA[3] := 10.0, [2,7].PID.DATA[4] := 10.0, [2,7].PID.DATA[5] := 0.02442002, [2,7].PID.DATA[6] := 1.0, [2,7].PID.DATA[7] := 4.3, [2,7].PID.DATA[8] := 2.0, [2,7].PID.DATA[9] := 0.2, [2,7].PID.DATA[10] := 0.3, [2,7].PID.DATA[11] := 2.0, [2,7].PID.DATA[12] := 0.2, [2,7].PID.DATA[13] := 0.3, [2,7].PID.DATA[15] := 1.0, [2,7].PID.DATA[16] := 1.0, [2,8].StableTimer.PRE := 15000, [2,8].PIDTimer.PRE := 250, [2,8].CycleTimer.PRE := 20000, [2,8].PID.CTL := 33555584, [2,8].PID.CA := 1, [2,8].PID.DVNA := 1, [2,8].PID.PVHA := 1, [2,8].PID.SP := 27.0, [2,8].PID.KP := 1.0, [2,8].PID.KI := 0.1, [2,8].PID.MAXS := 100.0, [2,8].PID.MAXO := 100.0, [2,8].PID.UPD := 0.25, [2,8].PID.PV := 18.2328, [2,8].PID.ERR := -8.767202, [2,8].PID.MAXI := 100.0, [2,8].PID.MAXCV := 100.0, [2,8].PID.MAXTIE := 100.0, [2,8].PID.DATA[0] := 8.767202, [2,8].PID.DATA[1] := 291.7248, [2,8].PID.DATA[2] := 18.2328, [2,8].PID.DATA[3] := -8.767202, [2,8].PID.DATA[4] := 27.0, [2,8].PID.DATA[5] := 1.0, [2,8].PID.DATA[6] := 1.0, [2,8].PID.DATA[7] := 4.0, [2,8].PID.DATA[8] := 1.0, [2,8].PID.DATA[9] := 0.1, [2,8].PID.DATA[11] := 1.0, [2,8].PID.DATA[12] := 0.1,
        [2,8].PID.DATA[15] := 1.0, [2,8].PID.DATA[16] := 1.0, [2,11].RampTimer.PRE := 100000, [2,11].StableTimer.PRE := 200, [2,11].PIDTimer.PRE := 250, [2,11].PIDTimer.ACC := 230, [2,11].PIDTimer.EN := 1, [2,11].PIDTimer.TT := 1, [2,11].PID.CTL := 67142528, [2,11].PID.SWM := 1, [2,11].PID.INI := 1, [2,11].PID.DVPA := 1, [2,11].PID.PVLA := 1, [2,11].PID.PVHA := 1, [2,11].PID.SP := 0.2, [2,11].PID.KP := 0.1, [2,11].PID.KI := 0.1, [2,11].PID.BIAS := 23.09767, [2,11].PID.DB := 0.001, [2,11].PID.MAXO := 100.0, [2,11].PID.UPD := 0.25, [2,11].PID.ERR := 0.2, [2,11].PID.MAXCV := 100.0, [2,11].PID.MAXTIE := 100.0, [2,11].PID.DATA[0] := -23.09816, [2,11].PID.DATA[3] := 0.2, [2,11].PID.DATA[4] := 0.2, [2,11].PID.DATA[5] := 0.02442002, [2,11].PID.DATA[6] := 1.0, [2,11].PID.DATA[7] := 4.0, [2,11].PID.DATA[8] := 0.1, [2,11].PID.DATA[9] := 0.1, [2,11].PID.DATA[11] := 0.1, [2,11].PID.DATA[12] := 0.1, [2,11].PID.DATA[15] := 1.0, [2,11].PID.DATA[16] := 1.0, [2,13].RampTimer.PRE := 3600000, [2,13].StableTimer.PRE := 2000, [2,13].PIDTimer.PRE := 10000, [2,13].PIDTimer.EN := 1, [2,13].PIDTimer.TT := 1, [2,13].PID.CTL := 305173120, [2,13].PID.PVT := 1, [2,13].PID.CA := 1, [2,13].PID.NOBC := 1, [2,13].PID.NOZC := 1, [2,13].PID.INI := 1, [2,13].PID.OLH := 1, [2,13].PID.DVPA := 1, [2,13].PID.PVHA := 1, [2,13].PID.KP := 0.2, [2,13].PID.KI := 0.08, [2,13].PID.MAXS := 100.0, [2,13].PID.DB := 1.0, [2,13].PID.SO := 100.0, [2,13].PID.MAXO := 100.0, [2,13].PID.UPD := 0.01, [2,13].PID.PV := 43.92523, [2,13].PID.ERR := 43.92523, [2,13].PID.OUT := 100.0,
        [2,13].PID.MAXI := 100.0, [2,13].PID.TIE := 2.442003, [2,13].PID.MAXCV := 100.0, [2,13].PID.MAXTIE := 4095.0, [2,13].PID.DATA[0] := 100.0, [2,13].PID.DATA[1] := 702.8037, [2,13].PID.DATA[2] := 43.92523, [2,13].PID.DATA[3] := 43.92523, [2,13].PID.DATA[5] := 1.0, [2,13].PID.DATA[6] := 1.0, [2,13].PID.DATA[7] := 0.16, [2,13].PID.DATA[8] := 0.2, [2,13].PID.DATA[9] := 0.08, [2,13].PID.DATA[11] := 0.2, [2,13].PID.DATA[12] := 0.08, [2,13].PID.DATA[15] := 1.0, [2,13].PID.DATA[16] := 0.02442002, [3,1].LoopCfg := 1, [3,1].DBOK := 1, [3,1].RampEnable := 1, [3,1].PIDEnable := 1, [3,1].RangeMax := 100.0, [3,1].RampRate := 0.5, [3,1].RampRateSave := 0.5, [3,1].RampTimer.PRE := 3600000, [3,1].PIDTimer.PRE := 250, [3,1].PIDTimer.EN := 1, [3,1].PIDTimer.TT := 1, [3,1].CycleTimer.PRE := 2000, [3,1].PID.CTL := 67108864, [3,1].PID.SWM := 1, [3,1].PID.MAXS := 25.0, [3,1].PID.MAXO := 100.0, [3,1].PID.MAXI := 25.0, [3,1].PID.MAXCV := 100.0, [3,1].PID.MAXTIE := 25.0, [3,1].PID.DATA[5] := 4.0, [3,1].PID.DATA[6] := 1.0, [3,1].PID.DATA[15] := 1.0, [3,1].PID.DATA[16] := 4.0, [3,1].Auto1Cfg := 1, [3,1].Auto2Cfg := 1, [3,1].Auto1PVCfg := 10, [3,1].Auto2PVCfg := 42, [3,1].Auto1RangeMax := 55.0, [3,2].LoopCfg := 1, [3,2].DBOK := 1, [3,2].RampEnable := 1, [3,2].PIDEnable := 1, [3,2].RangeMax := 100.0, [3,2].RampRate := 0.5, [3,2].RampRateSave := 0.5, [3,2].RampTimer.PRE := 3600000, [3,2].PIDTimer.PRE := 250, [3,2].PIDTimer.EN := 1, [3,2].PIDTimer.TT := 1, [3,2].CycleTimer.PRE := 2000, [3,2].PID.CTL := 67108864, [3,2].PID.SWM := 1, [3,2].PID.MAXO := 100.0,
        [3,2].PID.MAXCV := 100.0, [3,2].PID.MAXTIE := 100.0, [3,2].PID.DATA[5] := 0.024420025, [3,2].PID.DATA[6] := 1.0, [3,2].PID.DATA[15] := 1.0, [3,2].PID.DATA[16] := 1.0, [3,2].Auto1Cfg := 1, [3,2].Auto2Cfg := 1, [3,2].Auto1PVCfg := 12, [3,2].Auto2PVCfg := 43, [3,2].Auto1RangeMax := 30.0, [3,2].OutputAddress := 1, [3,3].LoopCfg := 1, [3,3].Enable := 1, [3,3].Manual := 1, [3,3].Status := 9, [3,3].RampEnable := 1, [3,3].PIDEnable := 1, [3,3].RangeMax := 100.0, [3,3].RampRate := 0.5, [3,3].RampRateSave := 0.5, [3,3].RampTimer.PRE := 3600000, [3,3].PIDTimer.PRE := 250, [3,3].PIDTimer.EN := 1, [3,3].PIDTimer.TT := 1, [3,3].CycleTimer.PRE := 2000, [3,3].PID.CTL := 67108864, [3,3].PID.SWM := 1, [3,3].PID.MAXS := 4095.0, [3,3].PID.MAXO := 100.0, [3,3].PID.MAXI := 4095.0, [3,3].PID.MAXCV := 100.0, [3,3].PID.MAXTIE := 100.0, [3,3].PID.DATA[5] := 0.024420025, [3,3].PID.DATA[6] := 1.0, [3,3].PID.DATA[15] := 1.0, [3,3].PID.DATA[16] := 1.0, [3,3].OutputAddress := 2, [4,0].RampTimer.PRE := 3600000, [4,0].StableTimer.PRE := 5000, [4,0].PIDTimer.PRE := 250, [4,0].PIDTimer.ACC := 100, [4,0].PIDTimer.EN := 1, [4,0].PIDTimer.TT := 1, [4,0].PID.CTL := 25199488, [4,0].PID.MO := 1, [4,0].PID.PE := 1, [4,0].PID.INI := 1, [4,0].PID.DVPA := 1, [4,0].PID.PVLA := 1, [4,0].PID.PVHA := 1, [4,0].PID.SP := 66.66666, [4,0].PID.KP := 0.5, [4,0].PID.KI := 0.1, [4,0].PID.MAXS := 200.0, [4,0].PID.SO := 10.0, [4,0].PID.MAXO := 100.0, [4,0].PID.MINO := 10.0, [4,0].PID.UPD := 0.25, [4,0].PID.ERR := 66.66666,
        [4,0].PID.OUT := 10.0, [4,0].PID.MAXI := 200.0, [4,0].PID.TIE := 10.0, [4,0].PID.MAXCV := 100.0, [4,0].PID.MAXTIE := 100.0, [4,0].PID.DATA[0] := -6.666666, [4,0].PID.DATA[3] := 66.66666, [4,0].PID.DATA[4] := 66.66666, [4,0].PID.DATA[5] := 0.5, [4,0].PID.DATA[6] := 1.0, [4,0].PID.DATA[7] := 4.0, [4,0].PID.DATA[8] := 0.5, [4,0].PID.DATA[9] := 0.1, [4,0].PID.DATA[11] := 0.5, [4,0].PID.DATA[12] := 0.08333334, [4,0].PID.DATA[15] := 1.0, [4,0].PID.DATA[16] := 1.0, [4,1].Tag := 'FIC01', [4,1].Desc := 'Prim. Feed Pump Control', [4,1].LoopCfg := 1, [4,1].ManualEGU := '%', [4,1].Auto1EGU := 'LPM', [4,1].Auto2EGU := 'cm/h', [4,1].Manual := 1, [4,1].DBOK := 1, [4,1].RampEnable := 1, [4,1].PIDEnable := 1, [4,1].ManualOSR := 1, [4,1].PVAuto2 := 2400.0, [4,1].RangeMax := 100.0, [4,1].RampRate := 5.0, [4,1].RampRateSave := 5.0, [4,1].Deadband := 5.0, [4,1].RampTimer.PRE := 3600000, [4,1].StableTimer.PRE := 10000, [4,1].StableTime := 10, [4,1].PIDTimer.PRE := 250, [4,1].PIDTimer.ACC := 107, [4,1].PIDTimer.EN := 1, [4,1].PIDTimer.TT := 1, [4,1].CycleTimer.PRE := 2000, [4,1].PID.CTL := 67143552, [4,1].PID.SWM := 1, [4,1].PID.INI := 1, [4,1].PID.DVNA := 1, [4,1].PID.DVPA := 1, [4,1].PID.PVLA := 1, [4,1].PID.PVHA := 1, [4,1].PID.KP := 0.7, [4,1].PID.KI := 1.4, [4,1].PID.KD := 0.013, [4,1].PID.MAXS := 22.0, [4,1].PID.DB := 0.001, [4,1].PID.MAXO := 100.0, [4,1].PID.UPD := 0.25, [4,1].PID.MAXI := 22.0, [4,1].PID.MAXCV := 100.0, [4,1].PID.MAXTIE := 22.0, [4,1].PID.DATA[5] := 4.5454545, [4,1].PID.DATA[6] := 1.0,
        [4,1].PID.DATA[7] := 4.013, [4,1].PID.DATA[8] := 0.7, [4,1].PID.DATA[9] := 1.4, [4,1].PID.DATA[10] := 0.013, [4,1].PID.DATA[11] := 0.7, [4,1].PID.DATA[12] := 1.4, [4,1].PID.DATA[13] := 0.013, [4,1].PID.DATA[15] := 1.0, [4,1].PID.DATA[16] := 4.5454545, [4,1].KP[0] := 700.0, [4,1].KI[0] := 1400.0, [4,1].KD[0] := 13.0, [4,1].Auto1Cfg := 1, [4,1].Auto2Cfg := 1, [4,1].Auto1PVCfg := 10, [4,1].Auto2PVCfg := 42, [4,1].Auto1RangeMax := 22.0, [4,1].Auto2RangeMax := 9999.0, [4,2].Tag := 'FIC02', [4,2].Desc := 'Sec. Feed Pump Control', [4,2].LoopCfg := 1, [4,2].ManualEGU := '%', [4,2].Auto1EGU := 'LPM', [4,2].Auto2EGU := 'cm/h', [4,2].Interlock := 1, [4,2].Manual := 1, [4,2].DBOK := 1, [4,2].RampEnable := 1, [4,2].PIDEnable := 1, [4,2].ManualOSR := 1, [4,2].PVAuto2 := 2400.0, [4,2].RangeMax := 100.0, [4,2].RampRate := 5.0, [4,2].RampRateSave := 5.0, [4,2].RampStart := 75.0, [4,2].Deadband := 5.0, [4,2].RampTimer.PRE := 3600000, [4,2].StableTimer.PRE := 10000, [4,2].StableTime := 10, [4,2].PIDTimer.PRE := 250, [4,2].PIDTimer.ACC := 108, [4,2].PIDTimer.EN := 1, [4,2].PIDTimer.TT := 1, [4,2].CycleTimer.PRE := 2000, [4,2].PID.CTL := 67143552, [4,2].PID.SWM := 1, [4,2].PID.INI := 1, [4,2].PID.DVNA := 1, [4,2].PID.DVPA := 1, [4,2].PID.PVLA := 1, [4,2].PID.PVHA := 1, [4,2].PID.KP := 0.7, [4,2].PID.KI := 1.4, [4,2].PID.KD := 0.013, [4,2].PID.MAXS := 22.0, [4,2].PID.DB := 0.001, [4,2].PID.MAXO := 100.0, [4,2].PID.UPD := 0.25, [4,2].PID.MAXI := 22.0, [4,2].PID.MAXCV := 100.0,
        [4,2].PID.MAXTIE := 100.0, [4,2].PID.DATA[5] := 4.5454545, [4,2].PID.DATA[6] := 1.0, [4,2].PID.DATA[7] := 4.013, [4,2].PID.DATA[8] := 0.7, [4,2].PID.DATA[9] := 1.4, [4,2].PID.DATA[10] := 0.013, [4,2].PID.DATA[11] := 0.7, [4,2].PID.DATA[12] := 1.4, [4,2].PID.DATA[13] := 0.013, [4,2].PID.DATA[15] := 1.0, [4,2].PID.DATA[16] := 1.0, [4,2].KP[0] := 700.0, [4,2].KI[0] := 1400.0, [4,2].KD[0] := 13.0, [4,2].DisOSR := 1, [4,2].Auto1Cfg := 1, [4,2].Auto2Cfg := 1, [4,2].Auto1PVCfg := 12, [4,2].Auto2PVCfg := 43, [4,2].Auto1RangeMax := 22.0, [4,2].Auto2RangeMax := 9999.0, [4,2].OutputAddress := 1, [4,3].Tag := 'PCV12', [4,3].Desc := 'Post Column PCV012 Control', [4,3].LoopCfg := 1, [4,3].ManualEGU := '%', [4,3].Enable := 1, [4,3].Manual := 1, [4,3].Stable := 1, [4,3].DBOK := 1, [4,3].Status := 3, [4,3].RampEnable := 1, [4,3].PIDEnable := 1, [4,3].ManualOSR := 1, [4,3].RangeMax := 100.0, [4,3].RampRate := 5.0, [4,3].RampRateSave := 5.0, [4,3].RampStart := 98.0, [4,3].RampTimer.PRE := 3600000, [4,3].StableTimer.PRE := 2300, [4,3].StableTimer.ACC := 2354, [4,3].StableTimer.EN := 1, [4,3].StableTimer.DN := 1, [4,3].PIDTimer.PRE := 250, [4,3].PIDTimer.ACC := 108, [4,3].PIDTimer.EN := 1, [4,3].PIDTimer.TT := 1, [4,3].CycleTimer.PRE := 2000, [4,3].PID.CTL := 201361280, [4,3].PID.DOE := 1, [4,3].PID.SWM := 1, [4,3].PID.INI := 1, [4,3].PID.DVNA := 1, [4,3].PID.DVPA := 1, [4,3].PID.PVLA := 1, [4,3].PID.PVHA := 1, [4,3].PID.KP := 0.001, [4,3].PID.KI := 0.001, [4,3].PID.BIAS := 30.796,
        [4,3].PID.MAXS := 4095.0, [4,3].PID.MAXO := 100.0, [4,3].PID.UPD := 0.01, [4,3].PID.MAXI := 4095.0, [4,3].PID.MAXCV := 100.0, [4,3].PID.MAXTIE := 100.0, [4,3].PID.DATA[0] := -30.796, [4,3].PID.DATA[5] := 0.024420025, [4,3].PID.DATA[6] := 1.0, [4,3].PID.DATA[7] := 0.16, [4,3].PID.DATA[8] := 0.001, [4,3].PID.DATA[9] := 0.001, [4,3].PID.DATA[11] := 0.001, [4,3].PID.DATA[12] := 0.001, [4,3].PID.DATA[15] := 1.0, [4,3].PID.DATA[16] := 1.0, [4,3].OutputAddress := 2, [4,4].Tag := 'PCV10', [4,4].Desc := 'Line Pump1 PCV010 Control', [4,4].ManualEGU := '%', [4,4].Manual := 1, [4,4].Status := 3, [4,4].RampEnable := 1, [4,4].PIDEnable := 1, [4,4].RangeMax := 100.0, [4,4].RampRate := 0.5, [4,4].RampRateSave := 0.5, [4,4].RampStart := 3.443, [4,4].RampTimer.PRE := 3600000, [4,4].StableTimer.PRE := 5000, [4,4].PIDTimer.PRE := 250, [4,4].CycleTimer.PRE := 2000, [4,4].PID.CTL := 35652992, [4,4].PID.CA := 1, [4,4].PID.NOBC := 1, [4,4].PID.DVNA := 1, [4,4].PID.PVLA := 1, [4,4].PID.PVHA := 1, [4,4].PID.SP := 19.6, [4,4].PID.KP := 0.1, [4,4].PID.KI := 0.3, [4,4].PID.MAXS := 150.0, [4,4].PID.MAXO := 100.0, [4,4].PID.UPD := 0.25, [4,4].PID.ERR := -19.6, [4,4].PID.MAXI := 150.0, [4,4].PID.MAXCV := 100.0, [4,4].PID.MAXTIE := 100.0, [4,4].PID.DATA[0] := 1.3066667, [4,4].PID.DATA[3] := -19.6, [4,4].PID.DATA[4] := 19.6, [4,4].PID.DATA[5] := 0.6666667, [4,4].PID.DATA[6] := 1.0, [4,4].PID.DATA[7] := 4.0, [4,4].PID.DATA[8] := 0.1, [4,4].PID.DATA[9] := 0.3, [4,4].PID.DATA[11] := 0.1, [4,4].PID.DATA[12] := 0.3, [4,4].PID.DATA[15] := 1.0, [4,4].PID.DATA[16] := 1.0,
        [4,4].OutputAddress := 2, [4,5].Tag := 'PCV11', [4,5].Desc := 'Line Pump2 PCV011 Control', [4,5].ManualEGU := '%', [4,5].Manual := 1, [4,5].Status := 3, [4,5].RampEnable := 1, [4,5].PIDEnable := 1, [4,5].RangeMax := 100.0, [4,5].RampRate := 0.5, [4,5].RampRateSave := 0.5, [4,5].RampStart := 4.417, [4,5].RampTimer.PRE := 3600000, [4,5].StableTimer.PRE := 1500, [4,5].PIDTimer.PRE := 250, [4,5].CycleTimer.PRE := 2000, [4,5].PID.CTL := 134218624, [4,5].PID.DOE := 1, [4,5].PID.DVPA := 1, [4,5].PID.PVLA := 1, [4,5].PID.PVHA := 1, [4,5].PID.SP := 350.0, [4,5].PID.KP := 40.0, [4,5].PID.KI := 0.5, [4,5].PID.BIAS := -847.4798, [4,5].PID.MAXS := 550.0, [4,5].PID.MAXO := 100.0, [4,5].PID.UPD := 0.25, [4,5].PID.ERR := 350.0, [4,5].PID.MAXI := 550.0, [4,5].PID.MAXCV := 100.0, [4,5].PID.MAXTIE := 100.0, [4,5].PID.DATA[0] := -1697.9749, [4,5].PID.DATA[1] := 1018.1818, [4,5].PID.DATA[3] := 350.0, [4,5].PID.DATA[4] := 350.0, [4,5].PID.DATA[5] := 0.18181819, [4,5].PID.DATA[6] := 1.0, [4,5].PID.DATA[7] := 4.0, [4,5].PID.DATA[8] := 40.0, [4,5].PID.DATA[9] := 0.5, [4,5].PID.DATA[11] := 40.0, [4,5].PID.DATA[12] := 0.5, [4,5].PID.DATA[15] := 1.0, [4,5].PID.DATA[16] := 1.0, [4,5].OutputAddress := 3, [4,6].StableTimer.PRE := 15000, [4,6].PIDTimer.EN := 1, [4,6].PIDTimer.TT := 1, [4,6].CycleTimer.PRE := 5000, [4,6].PID.CTL := 16810624, [4,6].PID.MO := 1, [4,6].PID.INI := 1, [4,6].PID.DVPA := 1, [4,6].PID.PVHA := 1, [4,6].PID.SP := 10.0, [4,6].PID.KP := 0.3, [4,6].PID.KI := 0.3, [4,6].PID.MAXS := 200.0, [4,6].PID.SO := 3.074094,
        [4,6].PID.MAXO := 100.0, [4,6].PID.UPD := 0.25, [4,6].PID.PV := 1.488363, [4,6].PID.ERR := 8.511638, [4,6].PID.OUT := 3.074094, [4,6].PID.MAXI := 200.0, [4,6].PID.TIE := 3.074094, [4,6].PID.MAXCV := 200.0, [4,6].PID.MAXTIE := 200.0, [4,6].PID.DATA[0] := 1.797348, [4,6].PID.DATA[1] := -11.9069, [4,6].PID.DATA[2] := 1.488363, [4,6].PID.DATA[3] := 8.511638, [4,6].PID.DATA[4] := 10.0, [4,6].PID.DATA[5] := 0.5, [4,6].PID.DATA[6] := 1.0, [4,6].PID.DATA[7] := 4.0, [4,6].PID.DATA[8] := 0.3, [4,6].PID.DATA[9] := 0.3, [4,6].PID.DATA[11] := 0.3, [4,6].PID.DATA[12] := 0.3, [4,6].PID.DATA[15] := 2.0, [4,6].PID.DATA[16] := 0.5, [4,7].StableTimer.PRE := 200, [4,7].PIDTimer.PRE := 250, [4,7].PIDTimer.EN := 1, [4,7].PIDTimer.TT := 1, [4,7].CycleTimer.PRE := 10000, [4,7].PID.CTL := 16810880, [4,7].PID.MO := 1, [4,7].PID.INI := 1, [4,7].PID.DVPA := 1, [4,7].PID.PVLA := 1, [4,7].PID.PVHA := 1, [4,7].PID.SP := 10.0, [4,7].PID.KP := 2.0, [4,7].PID.KI := 0.2, [4,7].PID.KD := 0.3, [4,7].PID.BIAS := 50.0, [4,7].PID.DB := 0.01, [4,7].PID.SO := 80.0, [4,7].PID.MAXO := 100.0, [4,7].PID.UPD := 0.25, [4,7].PID.ERR := 10.0, [4,7].PID.OUT := 80.0, [4,7].PID.TIE := 80.0, [4,7].PID.MAXCV := 100.0, [4,7].PID.MAXTIE := 100.0, [4,7].PID.DATA[0] := 29.511597, [4,7].PID.DATA[3] := 10.0, [4,7].PID.DATA[4] := 10.0, [4,7].PID.DATA[5] := 0.024420025, [4,7].PID.DATA[6] := 1.0, [4,7].PID.DATA[7] := 4.3, [4,7].PID.DATA[8] := 2.0, [4,7].PID.DATA[9] := 0.2, [4,7].PID.DATA[10] := 0.3, [4,7].PID.DATA[11] := 2.0, [4,7].PID.DATA[12] := 0.2, [4,7].PID.DATA[13] := 0.3,
        [4,7].PID.DATA[15] := 1.0, [4,7].PID.DATA[16] := 1.0, [4,8].StableTimer.PRE := 15000, [4,8].PIDTimer.PRE := 250, [4,8].CycleTimer.PRE := 20000, [4,8].PID.CTL := 33555584, [4,8].PID.CA := 1, [4,8].PID.DVNA := 1, [4,8].PID.PVHA := 1, [4,8].PID.SP := 27.0, [4,8].PID.KP := 1.0, [4,8].PID.KI := 0.1, [4,8].PID.MAXS := 100.0, [4,8].PID.MAXO := 100.0, [4,8].PID.UPD := 0.25, [4,8].PID.PV := 18.2328, [4,8].PID.ERR := -8.767202, [4,8].PID.MAXI := 100.0, [4,8].PID.MAXCV := 100.0, [4,8].PID.MAXTIE := 100.0, [4,8].PID.DATA[0] := 8.767202, [4,8].PID.DATA[1] := 291.7248, [4,8].PID.DATA[2] := 18.2328, [4,8].PID.DATA[3] := -8.767202, [4,8].PID.DATA[4] := 27.0, [4,8].PID.DATA[5] := 1.0, [4,8].PID.DATA[6] := 1.0, [4,8].PID.DATA[7] := 4.0, [4,8].PID.DATA[8] := 1.0, [4,8].PID.DATA[9] := 0.1, [4,8].PID.DATA[11] := 1.0, [4,8].PID.DATA[12] := 0.1, [4,8].PID.DATA[15] := 1.0, [4,8].PID.DATA[16] := 1.0, [4,11].RampTimer.PRE := 100000, [4,11].StableTimer.PRE := 200, [4,11].PIDTimer.PRE := 250, [4,11].PIDTimer.ACC := 230, [4,11].PIDTimer.EN := 1, [4,11].PIDTimer.TT := 1, [4,11].PID.CTL := 67142528, [4,11].PID.SWM := 1, [4,11].PID.INI := 1, [4,11].PID.DVPA := 1, [4,11].PID.PVLA := 1, [4,11].PID.PVHA := 1, [4,11].PID.SP := 0.20000005, [4,11].PID.KP := 0.1, [4,11].PID.KI := 0.1, [4,11].PID.BIAS := 23.09767, [4,11].PID.DB := 0.001, [4,11].PID.MAXO := 100.0, [4,11].PID.UPD := 0.25, [4,11].PID.ERR := 0.20000005, [4,11].PID.MAXCV := 100.0, [4,11].PID.MAXTIE := 100.0, [4,11].PID.DATA[0] := -23.098158, [4,11].PID.DATA[3] := 0.20000005, [4,11].PID.DATA[4] := 0.20000005, [4,11].PID.DATA[5] := 0.024420025,
        [4,11].PID.DATA[6] := 1.0, [4,11].PID.DATA[7] := 4.0, [4,11].PID.DATA[8] := 0.1, [4,11].PID.DATA[9] := 0.1, [4,11].PID.DATA[11] := 0.1, [4,11].PID.DATA[12] := 0.1, [4,11].PID.DATA[15] := 1.0, [4,11].PID.DATA[16] := 1.0, [4,13].RampTimer.PRE := 3600000, [4,13].StableTimer.PRE := 2000, [4,13].PIDTimer.PRE := 10000, [4,13].PIDTimer.EN := 1, [4,13].PIDTimer.TT := 1, [4,13].PID.CTL := 305173120, [4,13].PID.PVT := 1, [4,13].PID.CA := 1, [4,13].PID.NOBC := 1, [4,13].PID.NOZC := 1, [4,13].PID.INI := 1, [4,13].PID.OLH := 1, [4,13].PID.DVPA := 1, [4,13].PID.PVHA := 1, [4,13].PID.KP := 0.2, [4,13].PID.KI := 0.08, [4,13].PID.MAXS := 100.0, [4,13].PID.DB := 1.0, [4,13].PID.SO := 100.0, [4,13].PID.MAXO := 100.0, [4,13].PID.UPD := 0.01, [4,13].PID.PV := 43.925232, [4,13].PID.ERR := 43.925232, [4,13].PID.OUT := 100.0, [4,13].PID.MAXI := 100.0, [4,13].PID.TIE := 2.4420025, [4,13].PID.MAXCV := 100.0, [4,13].PID.MAXTIE := 4095.0, [4,13].PID.DATA[0] := 100.0, [4,13].PID.DATA[1] := 702.8037, [4,13].PID.DATA[2] := 43.925232, [4,13].PID.DATA[3] := 43.925232, [4,13].PID.DATA[5] := 1.0, [4,13].PID.DATA[6] := 1.0, [4,13].PID.DATA[7] := 0.16, [4,13].PID.DATA[8] := 0.2, [4,13].PID.DATA[9] := 0.08, [4,13].PID.DATA[11] := 0.2, [4,13].PID.DATA[12] := 0.08, [4,13].PID.DATA[15] := 1.0, [4,13].PID.DATA[16] := 0.024420025, [5,0].RampTimer.PRE := 3600000, [5,0].StableTimer.PRE := 5000, [5,0].PIDTimer.PRE := 250, [5,0].PIDTimer.ACC := 100, [5,0].PIDTimer.EN := 1, [5,0].PIDTimer.TT := 1, [5,0].PID.CTL := 25199488, [5,0].PID.MO := 1, [5,0].PID.PE := 1, [5,0].PID.INI := 1, [5,0].PID.DVPA := 1,
        [5,0].PID.PVLA := 1, [5,0].PID.PVHA := 1, [5,0].PID.SP := 66.66666, [5,0].PID.KP := 0.5, [5,0].PID.KI := 0.1, [5,0].PID.MAXS := 200.0, [5,0].PID.SO := 10.0, [5,0].PID.MAXO := 100.0, [5,0].PID.MINO := 10.0, [5,0].PID.UPD := 0.25, [5,0].PID.ERR := 66.66666, [5,0].PID.OUT := 10.0, [5,0].PID.MAXI := 200.0, [5,0].PID.TIE := 10.0, [5,0].PID.MAXCV := 100.0, [5,0].PID.MAXTIE := 100.0, [5,0].PID.DATA[0] := -6.666666, [5,0].PID.DATA[3] := 66.66666, [5,0].PID.DATA[4] := 66.66666, [5,0].PID.DATA[5] := 0.5, [5,0].PID.DATA[6] := 1.0, [5,0].PID.DATA[7] := 4.0, [5,0].PID.DATA[8] := 0.5, [5,0].PID.DATA[9] := 0.1, [5,0].PID.DATA[11] := 0.5, [5,0].PID.DATA[12] := 0.08333334, [5,0].PID.DATA[15] := 1.0, [5,0].PID.DATA[16] := 1.0, [5,1].Tag := 'FIC01', [5,1].Desc := 'Prim. Feed Pump Control', [5,1].LoopCfg := 1, [5,1].ManualEGU := '%', [5,1].Auto1EGU := 'LPM', [5,1].Auto2EGU := 'cm/h', [5,1].Manual := 1, [5,1].DBOK := 1, [5,1].RampEnable := 1, [5,1].PIDEnable := 1, [5,1].ManualOSR := 1, [5,1].PVAuto2 := 2400.0, [5,1].RangeMax := 100.0, [5,1].RampRate := 5.0, [5,1].RampRateSave := 5.0, [5,1].Deadband := 5.0, [5,1].RampTimer.PRE := 3600000, [5,1].StableTimer.PRE := 10000, [5,1].StableTime := 10, [5,1].PIDTimer.PRE := 250, [5,1].PIDTimer.EN := 1, [5,1].PIDTimer.TT := 1, [5,1].CycleTimer.PRE := 2000, [5,1].PID.CTL := 67143552, [5,1].PID.SWM := 1, [5,1].PID.INI := 1, [5,1].PID.DVNA := 1, [5,1].PID.DVPA := 1, [5,1].PID.PVLA := 1, [5,1].PID.PVHA := 1, [5,1].PID.KP := 0.7, [5,1].PID.KI := 1.4,
        [5,1].PID.KD := 0.013, [5,1].PID.DB := 0.001, [5,1].PID.MAXO := 100.0, [5,1].PID.UPD := 0.25, [5,1].PID.MAXCV := 100.0, [5,1].PID.DATA[5] := 0.024420025, [5,1].PID.DATA[6] := 1.0, [5,1].PID.DATA[7] := 4.013, [5,1].PID.DATA[8] := 0.7, [5,1].PID.DATA[9] := 1.4, [5,1].PID.DATA[10] := 0.013, [5,1].PID.DATA[11] := 0.7, [5,1].PID.DATA[12] := 1.4, [5,1].PID.DATA[13] := 0.013, [5,1].PID.DATA[15] := 1.0, [5,1].PID.DATA[16] := 1.0, [5,1].KP[0] := 700.0, [5,1].KI[0] := 1400.0, [5,1].KD[0] := 13.0, [5,1].Auto1Cfg := 1, [5,1].Auto2Cfg := 1, [5,1].Auto1PVCfg := 10, [5,1].Auto2PVCfg := 42, [5,1].Auto2RangeMax := 5.0, [5,2].Tag := 'FIC02', [5,2].Desc := 'Sec. Feed Pump Control', [5,2].LoopCfg := 1, [5,2].ManualEGU := '%', [5,2].Auto1EGU := 'LPM', [5,2].Auto2EGU := 'cm/h', [5,2].Interlock := 1, [5,2].Manual := 1, [5,2].DBOK := 1, [5,2].RampEnable := 1, [5,2].PIDEnable := 1, [5,2].ManualOSR := 1, [5,2].PVAuto2 := 2400.0, [5,2].RangeMax := 100.0, [5,2].RampRate := 5.0, [5,2].RampRateSave := 5.0, [5,2].RampStart := 75.0, [5,2].Deadband := 5.0, [5,2].RampTimer.PRE := 3600000, [5,2].StableTimer.PRE := 10000, [5,2].StableTime := 10, [5,2].PIDTimer.PRE := 250, [5,2].PIDTimer.EN := 1, [5,2].PIDTimer.TT := 1, [5,2].CycleTimer.PRE := 2000, [5,2].PID.CTL := 67143552, [5,2].PID.SWM := 1, [5,2].PID.INI := 1, [5,2].PID.DVNA := 1, [5,2].PID.DVPA := 1, [5,2].PID.PVLA := 1, [5,2].PID.PVHA := 1, [5,2].PID.KP := 0.7, [5,2].PID.KI := 1.4, [5,2].PID.KD := 0.013, [5,2].PID.MAXS := 50.0,
        [5,2].PID.DB := 0.001, [5,2].PID.MAXO := 100.0, [5,2].PID.UPD := 0.25, [5,2].PID.MAXI := 50.0, [5,2].PID.MAXCV := 100.0, [5,2].PID.MAXTIE := 100.0, [5,2].PID.DATA[5] := 2.0, [5,2].PID.DATA[6] := 1.0, [5,2].PID.DATA[7] := 4.013, [5,2].PID.DATA[8] := 0.7, [5,2].PID.DATA[9] := 1.4, [5,2].PID.DATA[10] := 0.013, [5,2].PID.DATA[11] := 0.7, [5,2].PID.DATA[12] := 1.4, [5,2].PID.DATA[13] := 0.013, [5,2].PID.DATA[15] := 1.0, [5,2].PID.DATA[16] := 1.0, [5,2].KP[0] := 700.0, [5,2].KI[0] := 1400.0, [5,2].KD[0] := 13.0, [5,2].DisOSR := 1, [5,2].Auto1Cfg := 1, [5,2].Auto2Cfg := 1, [5,2].Auto1PVCfg := 12, [5,2].Auto2PVCfg := 43, [5,2].Auto1RangeMax := 50.0, [5,2].Auto2RangeMax := 99999.0, [5,2].OutputAddress := 1, [5,3].Tag := 'PCV12', [5,3].Desc := 'Post Column PCV012 Control', [5,3].LoopCfg := 1, [5,3].ManualEGU := '%', [5,3].Enable := 1, [5,3].Manual := 1, [5,3].Stable := 1, [5,3].DBOK := 1, [5,3].Status := 3, [5,3].RampEnable := 1, [5,3].PIDEnable := 1, [5,3].ManualOSR := 1, [5,3].RangeMax := 100.0, [5,3].RampRate := 5.0, [5,3].RampRateSave := 5.0, [5,3].RampStart := 98.0, [5,3].RampTimer.PRE := 3600000, [5,3].StableTimer.PRE := 2300, [5,3].StableTimer.ACC := 2354, [5,3].StableTimer.EN := 1, [5,3].StableTimer.DN := 1, [5,3].PIDTimer.PRE := 250, [5,3].PIDTimer.EN := 1, [5,3].PIDTimer.TT := 1, [5,3].CycleTimer.PRE := 2000, [5,3].PID.CTL := 201361280, [5,3].PID.DOE := 1, [5,3].PID.SWM := 1, [5,3].PID.INI := 1, [5,3].PID.DVNA := 1, [5,3].PID.DVPA := 1, [5,3].PID.PVLA := 1,
        [5,3].PID.PVHA := 1, [5,3].PID.KP := 0.001, [5,3].PID.KI := 0.001, [5,3].PID.BIAS := 30.796, [5,3].PID.MAXS := 4095.0, [5,3].PID.MAXO := 100.0, [5,3].PID.UPD := 0.01, [5,3].PID.MAXI := 4095.0, [5,3].PID.MAXCV := 100.0, [5,3].PID.MAXTIE := 100.0, [5,3].PID.DATA[0] := -30.796, [5,3].PID.DATA[5] := 0.024420025, [5,3].PID.DATA[6] := 1.0, [5,3].PID.DATA[7] := 0.16, [5,3].PID.DATA[8] := 0.001, [5,3].PID.DATA[9] := 0.001, [5,3].PID.DATA[11] := 0.001, [5,3].PID.DATA[12] := 0.001, [5,3].PID.DATA[15] := 1.0, [5,3].PID.DATA[16] := 1.0, [5,3].OutputAddress := 2, [5,4].Tag := 'PCV10', [5,4].Desc := 'Line Pump1 PCV010 Control', [5,4].ManualEGU := '%', [5,4].Manual := 1, [5,4].Status := 3, [5,4].RampEnable := 1, [5,4].PIDEnable := 1, [5,4].RangeMax := 100.0, [5,4].RampRate := 0.5, [5,4].RampRateSave := 0.5, [5,4].RampStart := 3.443, [5,4].RampTimer.PRE := 3600000, [5,4].StableTimer.PRE := 5000, [5,4].PIDTimer.PRE := 250, [5,4].CycleTimer.PRE := 2000, [5,4].PID.CTL := 35652992, [5,4].PID.CA := 1, [5,4].PID.NOBC := 1, [5,4].PID.DVNA := 1, [5,4].PID.PVLA := 1, [5,4].PID.PVHA := 1, [5,4].PID.SP := 19.6, [5,4].PID.KP := 0.1, [5,4].PID.KI := 0.3, [5,4].PID.MAXS := 150.0, [5,4].PID.MAXO := 100.0, [5,4].PID.UPD := 0.25, [5,4].PID.ERR := -19.6, [5,4].PID.MAXI := 150.0, [5,4].PID.MAXCV := 100.0, [5,4].PID.MAXTIE := 100.0, [5,4].PID.DATA[0] := 1.3066667, [5,4].PID.DATA[3] := -19.6, [5,4].PID.DATA[4] := 19.6, [5,4].PID.DATA[5] := 0.6666667, [5,4].PID.DATA[6] := 1.0, [5,4].PID.DATA[7] := 4.0, [5,4].PID.DATA[8] := 0.1, [5,4].PID.DATA[9] := 0.3,
        [5,4].PID.DATA[11] := 0.1, [5,4].PID.DATA[12] := 0.3, [5,4].PID.DATA[15] := 1.0, [5,4].PID.DATA[16] := 1.0, [5,4].OutputAddress := 2, [5,5].Tag := 'PCV11', [5,5].Desc := 'Line Pump2 PCV011 Control', [5,5].ManualEGU := '%', [5,5].Manual := 1, [5,5].Status := 3, [5,5].RampEnable := 1, [5,5].PIDEnable := 1, [5,5].RangeMax := 100.0, [5,5].RampRate := 0.5, [5,5].RampRateSave := 0.5, [5,5].RampStart := 4.417, [5,5].RampTimer.PRE := 3600000, [5,5].StableTimer.PRE := 1500, [5,5].PIDTimer.PRE := 250, [5,5].CycleTimer.PRE := 2000, [5,5].PID.CTL := 134218624, [5,5].PID.DOE := 1, [5,5].PID.DVPA := 1, [5,5].PID.PVLA := 1, [5,5].PID.PVHA := 1, [5,5].PID.SP := 350.0, [5,5].PID.KP := 40.0, [5,5].PID.KI := 0.5, [5,5].PID.BIAS := -847.4798, [5,5].PID.MAXS := 550.0, [5,5].PID.MAXO := 100.0, [5,5].PID.UPD := 0.25, [5,5].PID.ERR := 350.0, [5,5].PID.MAXI := 550.0, [5,5].PID.MAXCV := 100.0, [5,5].PID.MAXTIE := 100.0, [5,5].PID.DATA[0] := -1697.9749, [5,5].PID.DATA[1] := 1018.1818, [5,5].PID.DATA[3] := 350.0, [5,5].PID.DATA[4] := 350.0, [5,5].PID.DATA[5] := 0.18181819, [5,5].PID.DATA[6] := 1.0, [5,5].PID.DATA[7] := 4.0, [5,5].PID.DATA[8] := 40.0, [5,5].PID.DATA[9] := 0.5, [5,5].PID.DATA[11] := 40.0, [5,5].PID.DATA[12] := 0.5, [5,5].PID.DATA[15] := 1.0, [5,5].PID.DATA[16] := 1.0, [5,5].OutputAddress := 3, [5,6].StableTimer.PRE := 15000, [5,6].PIDTimer.EN := 1, [5,6].PIDTimer.TT := 1, [5,6].CycleTimer.PRE := 5000, [5,6].PID.CTL := 16810624, [5,6].PID.MO := 1, [5,6].PID.INI := 1, [5,6].PID.DVPA := 1, [5,6].PID.PVHA := 1, [5,6].PID.SP := 10.0,
        [5,6].PID.KP := 0.3, [5,6].PID.KI := 0.3, [5,6].PID.MAXS := 200.0, [5,6].PID.SO := 3.074094, [5,6].PID.MAXO := 100.0, [5,6].PID.UPD := 0.25, [5,6].PID.PV := 1.488363, [5,6].PID.ERR := 8.511638, [5,6].PID.OUT := 3.074094, [5,6].PID.MAXI := 200.0, [5,6].PID.TIE := 3.074094, [5,6].PID.MAXCV := 200.0, [5,6].PID.MAXTIE := 200.0, [5,6].PID.DATA[0] := 1.797348, [5,6].PID.DATA[1] := -11.9069, [5,6].PID.DATA[2] := 1.488363, [5,6].PID.DATA[3] := 8.511638, [5,6].PID.DATA[4] := 10.0, [5,6].PID.DATA[5] := 0.5, [5,6].PID.DATA[6] := 1.0, [5,6].PID.DATA[7] := 4.0, [5,6].PID.DATA[8] := 0.3, [5,6].PID.DATA[9] := 0.3, [5,6].PID.DATA[11] := 0.3, [5,6].PID.DATA[12] := 0.3, [5,6].PID.DATA[15] := 2.0, [5,6].PID.DATA[16] := 0.5, [5,7].StableTimer.PRE := 200, [5,7].PIDTimer.PRE := 250, [5,7].PIDTimer.EN := 1, [5,7].PIDTimer.TT := 1, [5,7].CycleTimer.PRE := 10000, [5,7].PID.CTL := 16810880, [5,7].PID.MO := 1, [5,7].PID.INI := 1, [5,7].PID.DVPA := 1, [5,7].PID.PVLA := 1, [5,7].PID.PVHA := 1, [5,7].PID.SP := 10.0, [5,7].PID.KP := 2.0, [5,7].PID.KI := 0.2, [5,7].PID.KD := 0.3, [5,7].PID.BIAS := 50.0, [5,7].PID.DB := 0.01, [5,7].PID.SO := 80.0, [5,7].PID.MAXO := 100.0, [5,7].PID.UPD := 0.25, [5,7].PID.ERR := 10.0, [5,7].PID.OUT := 80.0, [5,7].PID.TIE := 80.0, [5,7].PID.MAXCV := 100.0, [5,7].PID.MAXTIE := 100.0, [5,7].PID.DATA[0] := 29.511597, [5,7].PID.DATA[3] := 10.0, [5,7].PID.DATA[4] := 10.0, [5,7].PID.DATA[5] := 0.024420025, [5,7].PID.DATA[6] := 1.0, [5,7].PID.DATA[7] := 4.3, [5,7].PID.DATA[8] := 2.0, [5,7].PID.DATA[9] := 0.2,
        [5,7].PID.DATA[10] := 0.3, [5,7].PID.DATA[11] := 2.0, [5,7].PID.DATA[12] := 0.2, [5,7].PID.DATA[13] := 0.3, [5,7].PID.DATA[15] := 1.0, [5,7].PID.DATA[16] := 1.0, [5,8].StableTimer.PRE := 15000, [5,8].PIDTimer.PRE := 250, [5,8].CycleTimer.PRE := 20000, [5,8].PID.CTL := 33555584, [5,8].PID.CA := 1, [5,8].PID.DVNA := 1, [5,8].PID.PVHA := 1, [5,8].PID.SP := 27.0, [5,8].PID.KP := 1.0, [5,8].PID.KI := 0.1, [5,8].PID.MAXS := 100.0, [5,8].PID.MAXO := 100.0, [5,8].PID.UPD := 0.25, [5,8].PID.PV := 18.2328, [5,8].PID.ERR := -8.767202, [5,8].PID.MAXI := 100.0, [5,8].PID.MAXCV := 100.0, [5,8].PID.MAXTIE := 100.0, [5,8].PID.DATA[0] := 8.767202, [5,8].PID.DATA[1] := 291.7248, [5,8].PID.DATA[2] := 18.2328, [5,8].PID.DATA[3] := -8.767202, [5,8].PID.DATA[4] := 27.0, [5,8].PID.DATA[5] := 1.0, [5,8].PID.DATA[6] := 1.0, [5,8].PID.DATA[7] := 4.0, [5,8].PID.DATA[8] := 1.0, [5,8].PID.DATA[9] := 0.1, [5,8].PID.DATA[11] := 1.0, [5,8].PID.DATA[12] := 0.1, [5,8].PID.DATA[15] := 1.0, [5,8].PID.DATA[16] := 1.0, [5,11].RampTimer.PRE := 100000, [5,11].StableTimer.PRE := 200, [5,11].PIDTimer.PRE := 250, [5,11].PIDTimer.ACC := 230, [5,11].PIDTimer.EN := 1, [5,11].PIDTimer.TT := 1, [5,11].PID.CTL := 67142528, [5,11].PID.SWM := 1, [5,11].PID.INI := 1, [5,11].PID.DVPA := 1, [5,11].PID.PVLA := 1, [5,11].PID.PVHA := 1, [5,11].PID.SP := 0.20000005, [5,11].PID.KP := 0.1, [5,11].PID.KI := 0.1, [5,11].PID.BIAS := 23.09767, [5,11].PID.DB := 0.001, [5,11].PID.MAXO := 100.0, [5,11].PID.UPD := 0.25, [5,11].PID.ERR := 0.20000005, [5,11].PID.MAXCV := 100.0, [5,11].PID.MAXTIE := 100.0,
        [5,11].PID.DATA[0] := -23.098158, [5,11].PID.DATA[3] := 0.20000005, [5,11].PID.DATA[4] := 0.20000005, [5,11].PID.DATA[5] := 0.024420025, [5,11].PID.DATA[6] := 1.0, [5,11].PID.DATA[7] := 4.0, [5,11].PID.DATA[8] := 0.1, [5,11].PID.DATA[9] := 0.1, [5,11].PID.DATA[11] := 0.1, [5,11].PID.DATA[12] := 0.1, [5,11].PID.DATA[15] := 1.0, [5,11].PID.DATA[16] := 1.0, [5,13].RampTimer.PRE := 3600000, [5,13].StableTimer.PRE := 2000, [5,13].PIDTimer.PRE := 10000, [5,13].PIDTimer.EN := 1, [5,13].PIDTimer.TT := 1, [5,13].PID.CTL := 305173120, [5,13].PID.PVT := 1, [5,13].PID.CA := 1, [5,13].PID.NOBC := 1, [5,13].PID.NOZC := 1, [5,13].PID.INI := 1, [5,13].PID.OLH := 1, [5,13].PID.DVPA := 1, [5,13].PID.PVHA := 1, [5,13].PID.KP := 0.2, [5,13].PID.KI := 0.08, [5,13].PID.MAXS := 100.0, [5,13].PID.DB := 1.0, [5,13].PID.SO := 100.0, [5,13].PID.MAXO := 100.0, [5,13].PID.UPD := 0.01, [5,13].PID.PV := 43.925232, [5,13].PID.ERR := 43.925232, [5,13].PID.OUT := 100.0, [5,13].PID.MAXI := 100.0, [5,13].PID.TIE := 2.4420025, [5,13].PID.MAXCV := 100.0, [5,13].PID.MAXTIE := 4095.0, [5,13].PID.DATA[0] := 100.0, [5,13].PID.DATA[1] := 702.8037, [5,13].PID.DATA[2] := 43.925232, [5,13].PID.DATA[3] := 43.925232, [5,13].PID.DATA[5] := 1.0, [5,13].PID.DATA[6] := 1.0, [5,13].PID.DATA[7] := 0.16, [5,13].PID.DATA[8] := 0.2, [5,13].PID.DATA[9] := 0.08, [5,13].PID.DATA[11] := 0.2, [5,13].PID.DATA[12] := 0.08, [5,13].PID.DATA[15] := 1.0, [5,13].PID.DATA[16] := 0.024420025);
   CPU_Scanning : BOOL := 1;   // System Scanning Flag
   CriteriaFlag : CriteriaFlag;   // Criteria Flag used in CCP Recipe
   DCS : DCS;
   DerivedData : DerivedData := (HOLDUP := 3.5, PI001_PSI := 0.0132753495, PI401_PSI := 0.33188373);   // Derived data (user input and calculated values)
   Diafiltration : Diafiltration := (Diaf_Init := 51.59, Diaf_Final_Volume := 10.0, Final_Diaf_Volum_DownTimer.PRE := 10000, Final_Diaf_Volum_DownTimer.ACC := 10089, Final_Diaf_Volum_DownTimer.EN := 1, Final_Diaf_Volum_DownTimer.DN := 1, Final_Diaf_Volum_UpTimer.PRE := 1000, LogDiafTimer.PRE := 3000);
   DigitalInput : BOOL[256] := ([0] := 1, [3] := 1, [4] := 1, [5] := 1, [8] := 1, [9] := 1, [10] := 1, [16] := 1, [17] := 1, [18] := 1, [19] := 1, [21] := 1, [22] := 1, [23] := 1, [24] := 1, [25] := 1, [100] := 1, [104] := 1, [106] := 1, [111] := 1, [131] := 1);   // Digital Input Array these bits are copied from Input cards.
   DigitalOutput : BOOL[256] := ([1] := 1, [34] := 1, [36] := 1, [37] := 1, [38] := 1, [39] := 1, [40] := 1, [41] := 1, [46] := 1, [180] := 1, [181] := 1);   // Digital Output Array these bits are sent to output cards.
        [4]   // Transfer Pump Run Command
        [7]   // Mixer Alarm Reset Command
        [17]   // spare
        [18]   // spare
        [19]   // spare
        [20]   // spare
        [21]   // spare
        [22]   // spare
        [23]   // spare
        [24]   // spare
        [25]   // spare
        [26]   // spare
        [27]   // spare
        [28]   // spare
        [29]   // spare
        [15]   // Connect Clamshell
        [12]   // Lock Clamshell
        [3]   // Feed Pump Run Command
        [11]   // Unlock Clamshell
        [0]   // Emergency Stop Acknowledge
        [9]   // Lock Door
        [1]   // Buzzer
        [10]   // Unlock Door
        [32]   // Valve XV001
        [33]   // Valve XV002
        [34]   // Valve XV003
        [35]   // Valve XV004
        [36]   // Valve XV005
        [37]   // Valve XV901
        [38]   // Valve XV102
        [39]   // Valve XV501
        [40]   // Valve XV502
        [41]   // Valve XV401
        [42]   // Valve XV402
        [43]   // Valve XV411
        [44]   // Valve XV421
        [45]   // Valve XV431
        [46]   // Valve XV441
        [47]   // Valve XV403
        [13]   // Unlock Clamshell in Door
        [30]   // spare
        [31]   // spare
        [48]   // Valve XV404
        [49]   // Valve XV405
        [50]   // Valve XV406
        [5]   // UV Auto zero
        [51]   // Valve XV006
        [52]   // Valve XV007
        [8]   // Feed Bag Tare
        [14]   // Lock Clamshell in Door
        [16]   // Disconnect Clamshell
        [2]   // Filtrate Bag Tare
        [6]   // Mixer Run Command
   DigitalPoint : DigitalPoint[150] := ([0].Tag := 'PSL602', [0].CurrentValue := 1, [0].Mimic := 1, [0].DelayTimer.PRE := 2000, [0].DelayTimerSP := 2, [0].Priority := 1, [0].EnableCfg := 1, [0].ActiveStateCFg := 1, [0].RealInputCfg := 1, [0].AlarmCfg := 1, [0].OverrideCfg := 1, [0].PriorityCfg := 1, [1].Tag := 'XS001', [1].AlarmCurrentValue := 1, [1].Override := 1, [1].Condition2 := 1, [1].DelayTimer.PRE := 1000, [1].DelayTimer.ACC := 1005, [1].DelayTimer.EN := 1, [1].DelayTimer.DN := 1, [1].DelayTimerSP := 1, [1].Priority := 1, [1].EnableCfg := 1, [1].ActiveStateCFg := 1, [1].RealInputCfg := 1, [1].InputAddressCfg := 1, [1].AlarmCfg := 1, [1].OverrideCfg := 1, [2].Tag := 'XS006', [2].DelayTimer.PRE := 1000, [2].DelayTimerSP := 1, [2].EnableCfg := 1, [2].ActiveStateCFg := 1, [2].RealInputCfg := 1, [2].InputAddressCfg := 2, [3].Tag := 'ES001', [3].CurrentValue := 1, [3].Mimic := 1, [3].Priority := 1, [3].EnableCfg := 1, [3].ActiveStateCFg := 1, [3].RealInputCfg := 1, [3].InputAddressCfg := 3, [3].AlarmCfg := 1, [4].Tag := 'PSH001', [4].CurrentValue := 1, [4].Override := 1, [4].Mimic := 1, [4].Priority := 1, [4].EnableCfg := 1, [4].ActiveStateCFg := 1, [4].RealInputCfg := 1, [4].InputAddressCfg := 4, [4].AlarmCfg := 1, [4].OverrideCfg := 1, [5].Tag := 'PSH401', [5].CurrentValue := 1, [5].Override := 1, [5].Mimic := 1, [5].Priority := 1,
        [5].EnableCfg := 1, [5].ActiveStateCFg := 1, [5].RealInputCfg := 1, [5].InputAddressCfg := 5, [5].AlarmCfg := 1, [5].OverrideCfg := 1, [6].Tag := 'XS002', [6].DelayTimer.PRE := 1000, [6].DelayTimerSP := 1, [6].EnableCfg := 1, [6].ActiveStateCFg := 1, [6].RealInputCfg := 1, [6].InputAddressCfg := 6, [7].Tag := 'XS003', [7].DelayTimer.PRE := 1000, [7].DelayTimerSP := 1, [7].EnableCfg := 1, [7].ActiveStateCFg := 1, [7].RealInputCfg := 1, [7].InputAddressCfg := 7, [8].Tag := 'SIC001DF', [8].CurrentValue := 1, [8].Mimic := 1, [8].DelayTimer.PRE := 1000, [8].DelayTimerSP := 1, [8].EnableCfg := 1, [8].ActiveStateCFg := 1, [8].RealInputCfg := 1, [8].InputAddressCfg := 8, [8].AlarmCfg := 1, [8].OverrideCfg := 1, [8].PriorityCfg := 1, [9].Tag := 'SIC002DF', [9].CurrentValue := 1, [9].Mimic := 1, [9].DelayTimer.PRE := 1000, [9].DelayTimerSP := 1, [9].Priority := 1, [9].EnableCfg := 1, [9].ActiveStateCFg := 1, [9].RealInputCfg := 1, [9].InputAddressCfg := 9, [9].AlarmCfg := 1, [9].OverrideCfg := 1, [9].PriorityCfg := 1, [10].Tag := 'PSL603', [10].CurrentValue := 1, [10].Mimic := 1, [10].DelayTimer.PRE := 2000, [10].DelayTimerSP := 2, [10].Priority := 1, [10].EnableCfg := 1, [10].ActiveStateCFg := 1, [10].RealInputCfg := 1, [10].InputAddressCfg := 10, [10].AlarmCfg := 1, [10].OverrideCfg := 1, [10].PriorityCfg := 1, [11].Tag := 'XS011', [11].DelayTimer.PRE := 1000,
